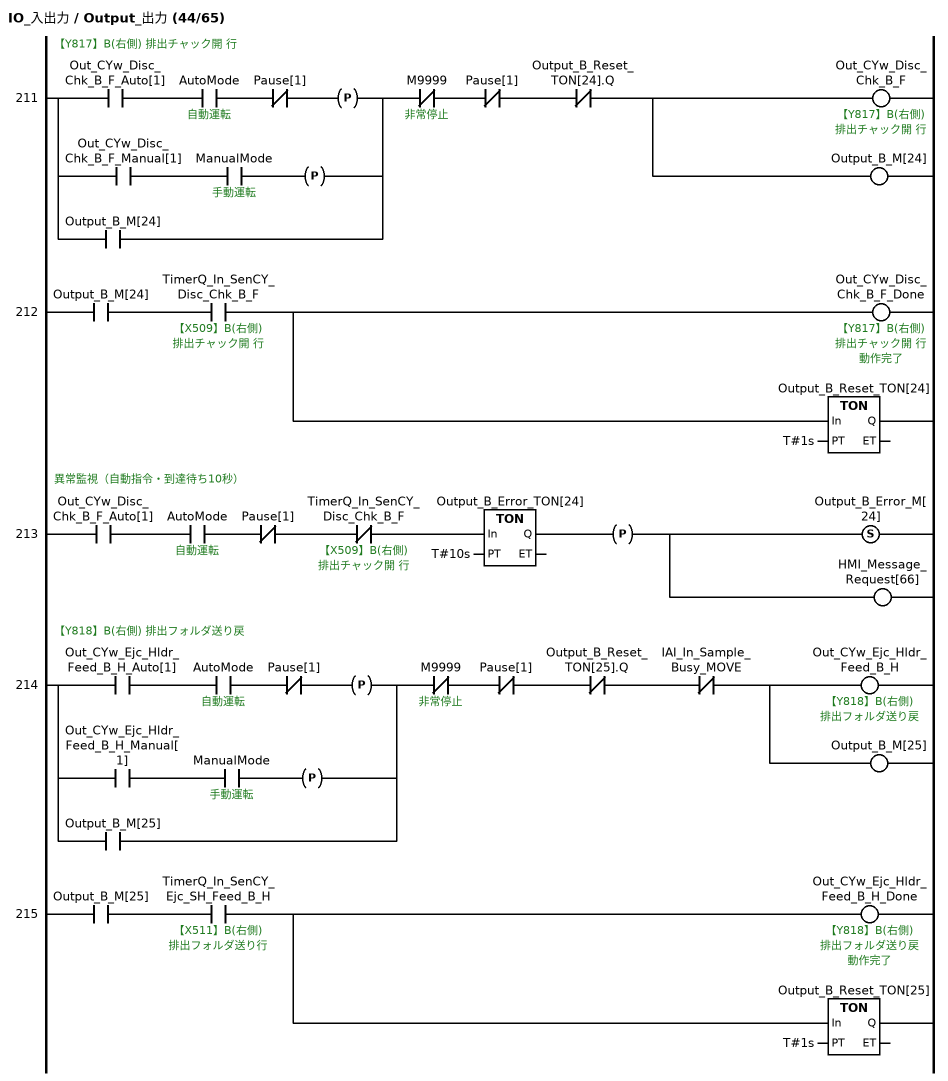
(* [picture p187: IO_入出力 / Output_出力, rungs 211-215] *)
(* Rung 211: 【Y817】B(右側) 排出チャック開 行 *)
_e309(CLK := Out_CYw_Disc_Chk_B_F_Auto[1] AND AutoMode AND NOT Pause[1]);
_e310(CLK := Out_CYw_Disc_Chk_B_F_Manual[1] AND ManualMode);
_p311 := (_e309.Q OR _e310.Q OR Output_B_M[24]) AND NOT M9999 AND NOT Pause[1] AND NOT Output_B_Reset_TON[24].Q;
Out_CYw_Disc_Chk_B_F := _p311;
Output_B_M[24] := _p311;
(* Rung 212 *)
Out_CYw_Disc_Chk_B_F_Done := Output_B_M[24] AND TimerQ_In_SenCY_Disc_Chk_B_F;
Output_B_Reset_TON[24](In := Output_B_M[24] AND TimerQ_In_SenCY_Disc_Chk_B_F, PT := T#1s);
(* Rung 213: 異常監視（自動指令・到達待ち10秒） *)
Output_B_Error_TON[24](In := Out_CYw_Disc_Chk_B_F_Auto[1] AND AutoMode AND NOT Pause[1] AND NOT TimerQ_In_SenCY_Disc_Chk_B_F, PT := T#10s);
_e312(CLK := Output_B_Error_TON[24].Q);
IF _e312.Q THEN Output_B_Error_M[24] := TRUE; END_IF;
HMI_Message_Request[66] := _e312.Q;
(* Rung 214: 【Y818】B(右側) 排出フォルダ送り戻 *)
_e313(CLK := Out_CYw_Ejc_Hldr_Feed_B_H_Auto[1] AND AutoMode AND NOT Pause[1]);
_e314(CLK := Out_CYw_Ejc_Hldr_Feed_B_H_Manual[1] AND ManualMode);
_p315 := (_e313.Q OR _e314.Q OR Output_B_M[25]) AND NOT M9999 AND NOT Pause[1] AND NOT Output_B_Reset_TON[25].Q AND NOT IAI_In_Sample_Busy_MOVE;
Out_CYw_Ejc_Hldr_Feed_B_H := _p315;
Output_B_M[25] := _p315;
(* Rung 215 *)
_p316 := Output_B_M[25] AND TimerQ_In_SenCY_Ejc_SH_Feed_B_H;
Out_CYw_Ejc_Hldr_Feed_B_H_Done := _p316;
Output_B_Reset_TON[25](In := _p316, PT := T#1s);

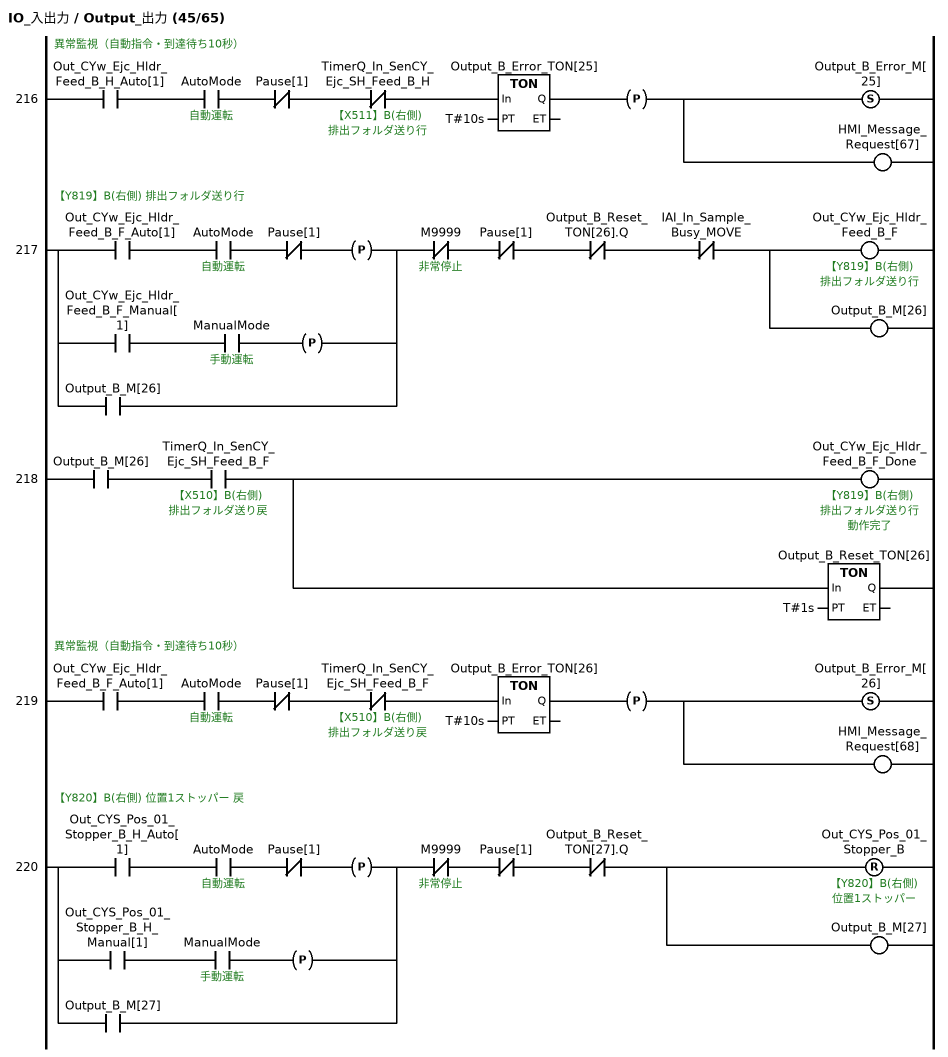
(* Rung 216: 異常監視（自動指令・到達待ち10秒） *)
Output_B_Error_TON[25](In := Out_CYw_Ejc_Hldr_Feed_B_H_Auto[1] AND AutoMode AND NOT Pause[1] AND NOT TimerQ_In_SenCY_Ejc_SH_Feed_B_H, PT := T#10s);
_e317(CLK := Output_B_Error_TON[25].Q);
IF _e317.Q THEN Output_B_Error_M[25] := TRUE; END_IF;
HMI_Message_Request[67] := _e317.Q;
(* Rung 217: 【Y819】B(右側) 排出フォルダ送り行 *)
_e318(CLK := Out_CYw_Ejc_Hldr_Feed_B_F_Auto[1] AND AutoMode AND NOT Pause[1]);
_e319(CLK := Out_CYw_Ejc_Hldr_Feed_B_F_Manual[1] AND ManualMode);
_p320 := (_e318.Q OR _e319.Q OR Output_B_M[26]) AND NOT M9999 AND NOT Pause[1] AND NOT Output_B_Reset_TON[26].Q AND NOT IAI_In_Sample_Busy_MOVE;
Out_CYw_Ejc_Hldr_Feed_B_F := _p320;
Output_B_M[26] := _p320;
(* Rung 218 *)
_p321 := Output_B_M[26] AND TimerQ_In_SenCY_Ejc_SH_Feed_B_F;
Out_CYw_Ejc_Hldr_Feed_B_F_Done := _p321;
Output_B_Reset_TON[26](In := _p321, PT := T#1s);
(* Rung 219: 異常監視（自動指令・到達待ち10秒） *)
Output_B_Error_TON[26](In := Out_CYw_Ejc_Hldr_Feed_B_F_Auto[1] AND AutoMode AND NOT Pause[1] AND NOT TimerQ_In_SenCY_Ejc_SH_Feed_B_F, PT := T#10s);
_e322(CLK := Output_B_Error_TON[26].Q);
IF _e322.Q THEN Output_B_Error_M[26] := TRUE; END_IF;
HMI_Message_Request[68] := _e322.Q;
(* Rung 220: 【Y820】B(右側) 位置1ストッパー 戻 *)
_e323(CLK := Out_CYS_Pos_01_Stopper_B_H_Auto[1] AND AutoMode AND NOT Pause[1]);
_e324(CLK := Out_CYS_Pos_01_Stopper_B_H_Manual[1] AND ManualMode);
_p325 := (_e323.Q OR _e324.Q OR Output_B_M[27]) AND NOT M9999 AND NOT Pause[1] AND NOT Output_B_Reset_TON[27].Q;
IF _p325 THEN Out_CYS_Pos_01_Stopper_B := FALSE; END_IF;
Output_B_M[27] := _p325;

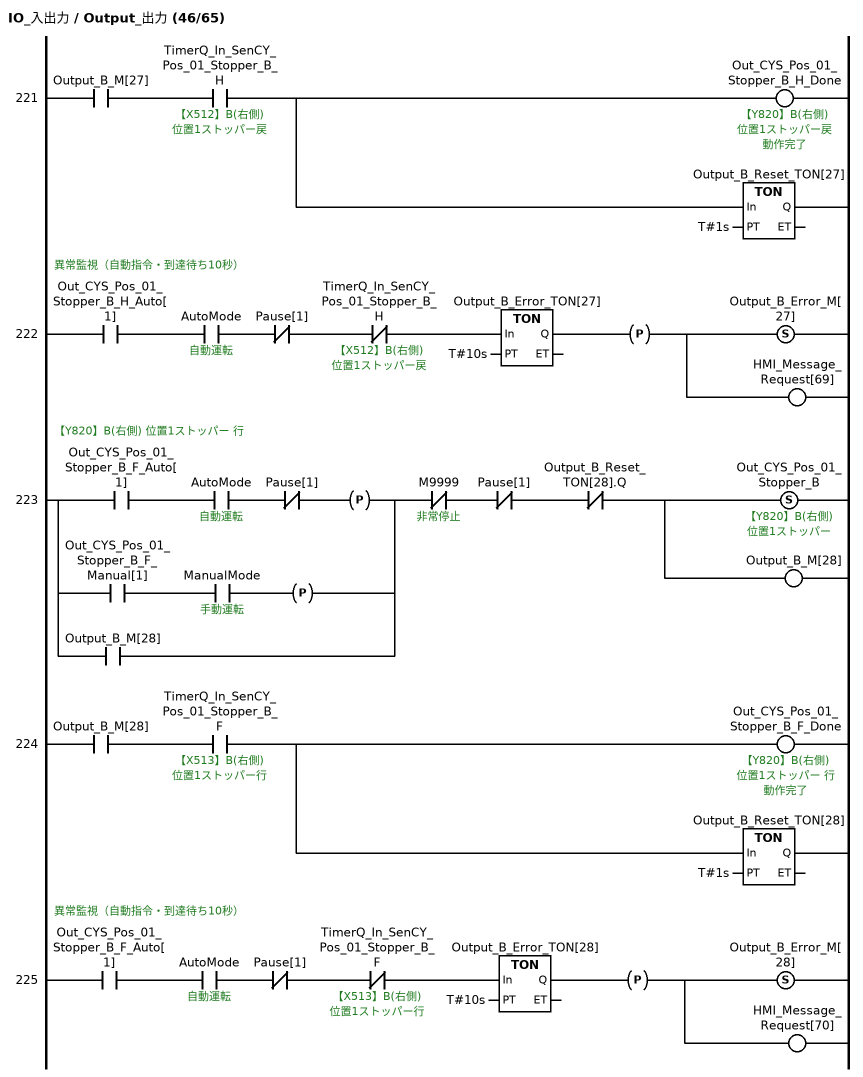
(* Rung 221 *)
_p326 := Output_B_M[27] AND TimerQ_In_SenCY_Pos_01_Stopper_B_H;
Out_CYS_Pos_01_Stopper_B_H_Done := _p326;
Output_B_Reset_TON[27](In := _p326, PT := T#1s);
(* Rung 222: 異常監視（自動指令・到達待ち10秒） *)
Output_B_Error_TON[27](In := Out_CYS_Pos_01_Stopper_B_H_Auto[1] AND AutoMode AND NOT Pause[1] AND NOT TimerQ_In_SenCY_Pos_01_Stopper_B_H, PT := T#10s);
_e327(CLK := Output_B_Error_TON[27].Q);
IF _e327.Q THEN Output_B_Error_M[27] := TRUE; END_IF;
HMI_Message_Request[69] := _e327.Q;
(* Rung 223: 【Y820】B(右側) 位置1ストッパー 行 *)
_e328(CLK := Out_CYS_Pos_01_Stopper_B_F_Auto[1] AND AutoMode AND NOT Pause[1]);
_e329(CLK := Out_CYS_Pos_01_Stopper_B_F_Manual[1] AND ManualMode);
_p330 := (_e328.Q OR _e329.Q OR Output_B_M[28]) AND NOT M9999 AND NOT Pause[1] AND NOT Output_B_Reset_TON[28].Q;
IF _p330 THEN Out_CYS_Pos_01_Stopper_B := TRUE; END_IF;
Output_B_M[28] := _p330;
(* Rung 224 *)
_p331 := Output_B_M[28] AND TimerQ_In_SenCY_Pos_01_Stopper_B_F;
Out_CYS_Pos_01_Stopper_B_F_Done := _p331;
Output_B_Reset_TON[28](In := _p331, PT := T#1s);
(* Rung 225: 異常監視（自動指令・到達待ち10秒） *)
Output_B_Error_TON[28](In := Out_CYS_Pos_01_Stopper_B_F_Auto[1] AND AutoMode AND NOT Pause[1] AND NOT TimerQ_In_SenCY_Pos_01_Stopper_B_F, PT := T#10s);
_e332(CLK := Output_B_Error_TON[28].Q);
IF _e332.Q THEN Output_B_Error_M[28] := TRUE; END_IF;
HMI_Message_Request[70] := _e332.Q;

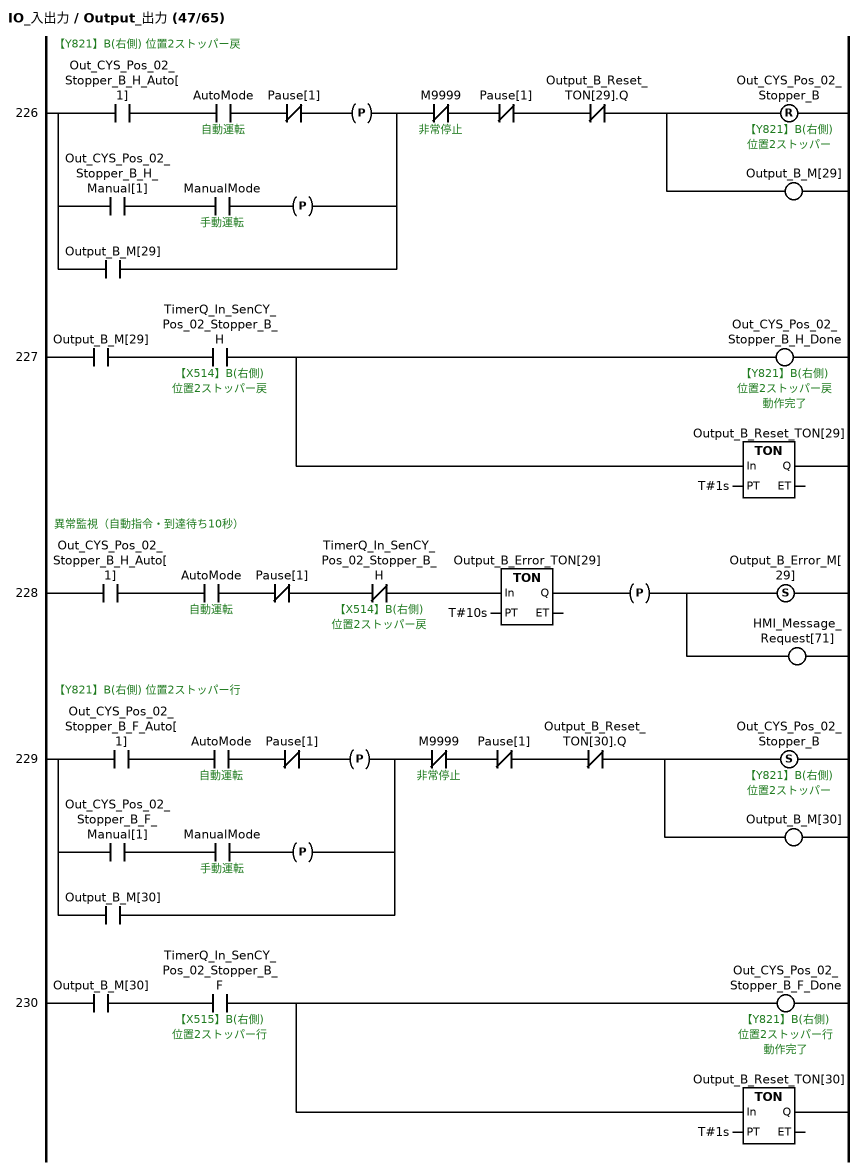
(* Rung 226: 【Y821】B(右側) 位置2ストッパー戻 *)
_e333(CLK := Out_CYS_Pos_02_Stopper_B_H_Auto[1] AND AutoMode AND NOT Pause[1]);
_e334(CLK := Out_CYS_Pos_02_Stopper_B_H_Manual[1] AND ManualMode);
_p335 := (_e333.Q OR _e334.Q OR Output_B_M[29]) AND NOT M9999 AND NOT Pause[1] AND NOT Output_B_Reset_TON[29].Q;
IF _p335 THEN Out_CYS_Pos_02_Stopper_B := FALSE; END_IF;
Output_B_M[29] := _p335;
(* Rung 227 *)
_p336 := Output_B_M[29] AND TimerQ_In_SenCY_Pos_02_Stopper_B_H;
Out_CYS_Pos_02_Stopper_B_H_Done := _p336;
Output_B_Reset_TON[29](In := _p336, PT := T#1s);
(* Rung 228: 異常監視（自動指令・到達待ち10秒） *)
Output_B_Error_TON[29](In := Out_CYS_Pos_02_Stopper_B_H_Auto[1] AND AutoMode AND NOT Pause[1] AND NOT TimerQ_In_SenCY_Pos_02_Stopper_B_H, PT := T#10s);
_e337(CLK := Output_B_Error_TON[29].Q);
IF _e337.Q THEN Output_B_Error_M[29] := TRUE; END_IF;
HMI_Message_Request[71] := _e337.Q;
(* Rung 229: 【Y821】B(右側) 位置2ストッパー行 *)
_e338(CLK := Out_CYS_Pos_02_Stopper_B_F_Auto[1] AND AutoMode AND NOT Pause[1]);
_e339(CLK := Out_CYS_Pos_02_Stopper_B_F_Manual[1] AND ManualMode);
_p340 := (_e338.Q OR _e339.Q OR Output_B_M[30]) AND NOT M9999 AND NOT Pause[1] AND NOT Output_B_Reset_TON[30].Q;
IF _p340 THEN Out_CYS_Pos_02_Stopper_B := TRUE; END_IF;
Output_B_M[30] := _p340;
(* Rung 230 *)
_p341 := Output_B_M[30] AND TimerQ_In_SenCY_Pos_02_Stopper_B_F;
Out_CYS_Pos_02_Stopper_B_F_Done := _p341;
Output_B_Reset_TON[30](In := _p341, PT := T#1s);

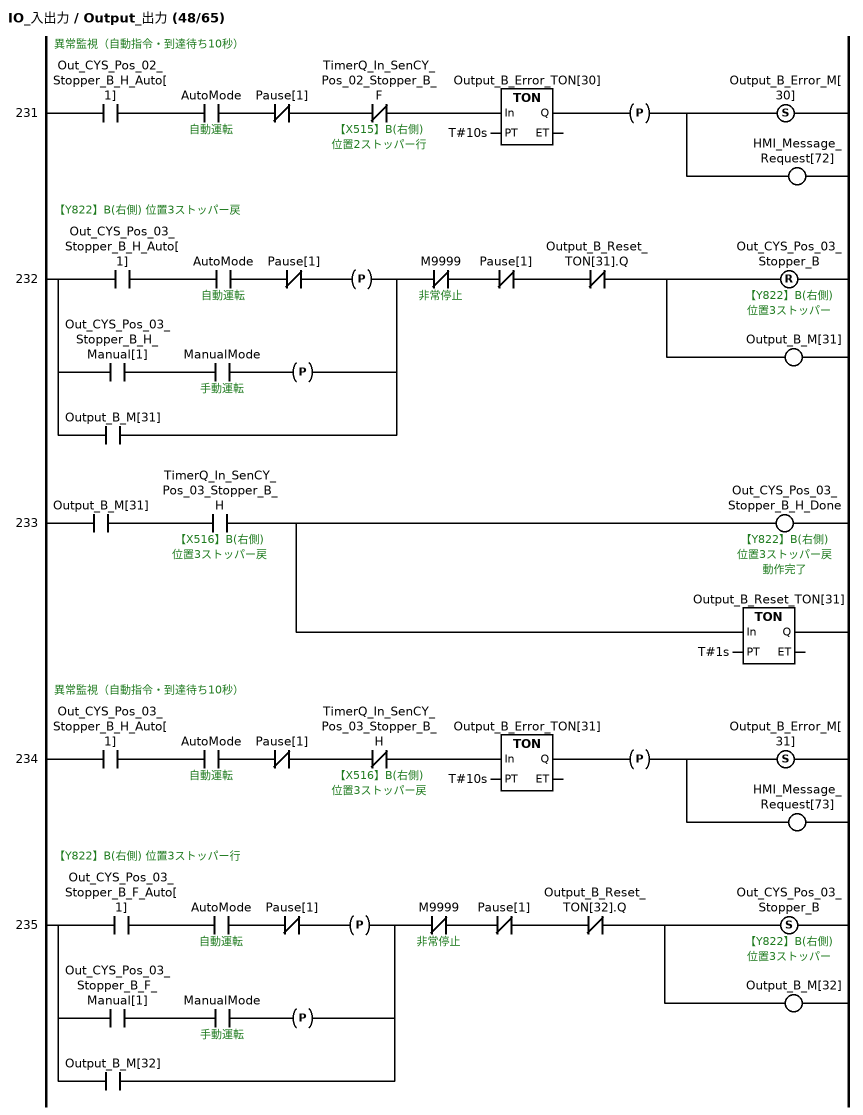
(* Rung 231: 異常監視（自動指令・到達待ち10秒） *)
Output_B_Error_TON[30](In := Out_CYS_Pos_02_Stopper_B_H_Auto[1] AND AutoMode AND NOT Pause[1] AND NOT TimerQ_In_SenCY_Pos_02_Stopper_B_F, PT := T#10s);
_e342(CLK := Output_B_Error_TON[30].Q);
IF _e342.Q THEN Output_B_Error_M[30] := TRUE; END_IF;
HMI_Message_Request[72] := _e342.Q;
(* Rung 232: 【Y822】B(右側) 位置3ストッパー戻 *)
_e343(CLK := Out_CYS_Pos_03_Stopper_B_H_Auto[1] AND AutoMode AND NOT Pause[1]);
_e344(CLK := Out_CYS_Pos_03_Stopper_B_H_Manual[1] AND ManualMode);
_p345 := (_e343.Q OR _e344.Q OR Output_B_M[31]) AND NOT M9999 AND NOT Pause[1] AND NOT Output_B_Reset_TON[31].Q;
IF _p345 THEN Out_CYS_Pos_03_Stopper_B := FALSE; END_IF;
Output_B_M[31] := _p345;
(* Rung 233 *)
_p346 := Output_B_M[31] AND TimerQ_In_SenCY_Pos_03_Stopper_B_H;
Out_CYS_Pos_03_Stopper_B_H_Done := _p346;
Output_B_Reset_TON[31](In := _p346, PT := T#1s);
(* Rung 234: 異常監視（自動指令・到達待ち10秒） *)
Output_B_Error_TON[31](In := Out_CYS_Pos_03_Stopper_B_H_Auto[1] AND AutoMode AND NOT Pause[1] AND NOT TimerQ_In_SenCY_Pos_03_Stopper_B_H, PT := T#10s);
_e347(CLK := Output_B_Error_TON[31].Q);
IF _e347.Q THEN Output_B_Error_M[31] := TRUE; END_IF;
HMI_Message_Request[73] := _e347.Q;
(* Rung 235: 【Y822】B(右側) 位置3ストッパー行 *)
_e348(CLK := Out_CYS_Pos_03_Stopper_B_F_Auto[1] AND AutoMode AND NOT Pause[1]);
_e349(CLK := Out_CYS_Pos_03_Stopper_B_F_Manual[1] AND ManualMode);
_p350 := (_e348.Q OR _e349.Q OR Output_B_M[32]) AND NOT M9999 AND NOT Pause[1] AND NOT Output_B_Reset_TON[32].Q;
IF _p350 THEN Out_CYS_Pos_03_Stopper_B := TRUE; END_IF;
Output_B_M[32] := _p350;

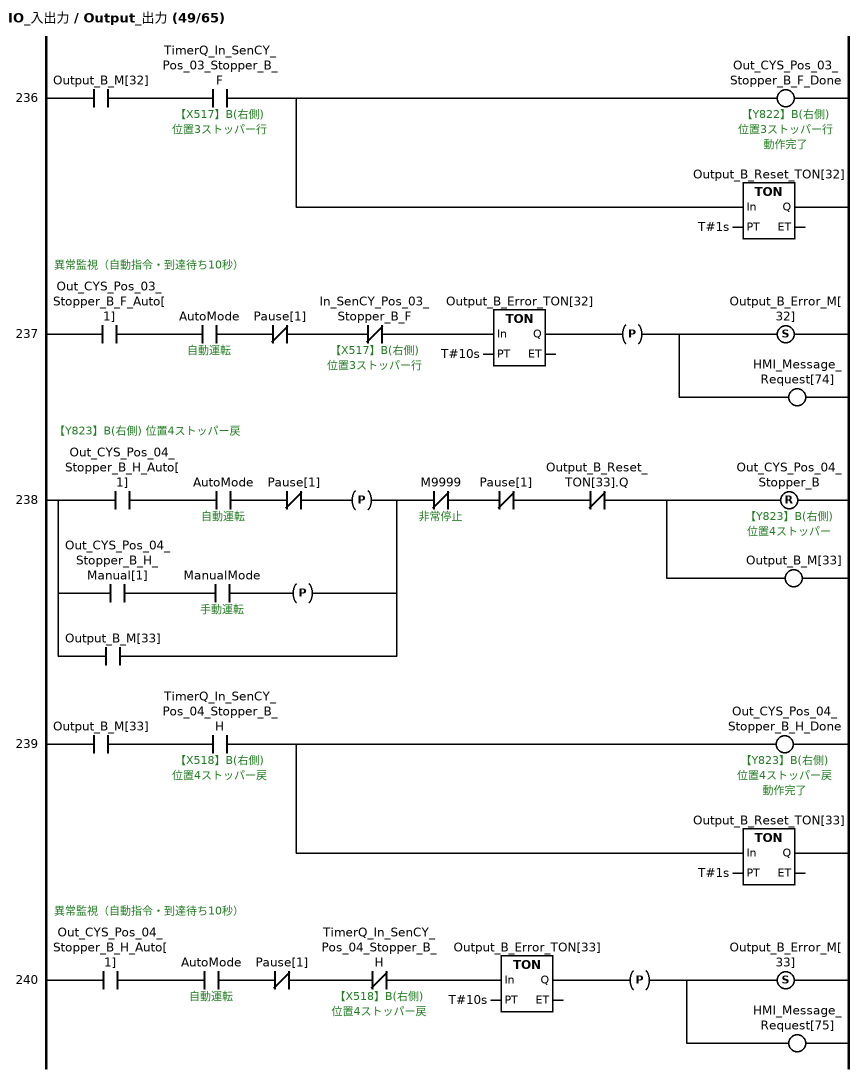
(* Rung 236 *)
_p351 := Output_B_M[32] AND TimerQ_In_SenCY_Pos_03_Stopper_B_F;
Out_CYS_Pos_03_Stopper_B_F_Done := _p351;
Output_B_Reset_TON[32](In := _p351, PT := T#1s);
(* Rung 237: 異常監視（自動指令・到達待ち10秒） *)
Output_B_Error_TON[32](In := Out_CYS_Pos_03_Stopper_B_F_Auto[1] AND AutoMode AND NOT Pause[1] AND NOT In_SenCY_Pos_03_Stopper_B_F, PT := T#10s);
_e352(CLK := Output_B_Error_TON[32].Q);
IF _e352.Q THEN Output_B_Error_M[32] := TRUE; END_IF;
HMI_Message_Request[74] := _e352.Q;
(* Rung 238: 【Y823】B(右側) 位置4ストッパー戻 *)
_e353(CLK := Out_CYS_Pos_04_Stopper_B_H_Auto[1] AND AutoMode AND NOT Pause[1]);
_e354(CLK := Out_CYS_Pos_04_Stopper_B_H_Manual[1] AND ManualMode);
_p355 := (_e353.Q OR _e354.Q OR Output_B_M[33]) AND NOT M9999 AND NOT Pause[1] AND NOT Output_B_Reset_TON[33].Q;
IF _p355 THEN Out_CYS_Pos_04_Stopper_B := FALSE; END_IF;
Output_B_M[33] := _p355;
(* Rung 239 *)
_p356 := Output_B_M[33] AND TimerQ_In_SenCY_Pos_04_Stopper_B_H;
Out_CYS_Pos_04_Stopper_B_H_Done := _p356;
Output_B_Reset_TON[33](In := _p356, PT := T#1s);
(* Rung 240: 異常監視（自動指令・到達待ち10秒） *)
Output_B_Error_TON[33](In := Out_CYS_Pos_04_Stopper_B_H_Auto[1] AND AutoMode AND NOT Pause[1] AND NOT TimerQ_In_SenCY_Pos_04_Stopper_B_H, PT := T#10s);
_e357(CLK := Output_B_Error_TON[33].Q);
IF _e357.Q THEN Output_B_Error_M[33] := TRUE; END_IF;
HMI_Message_Request[75] := _e357.Q;

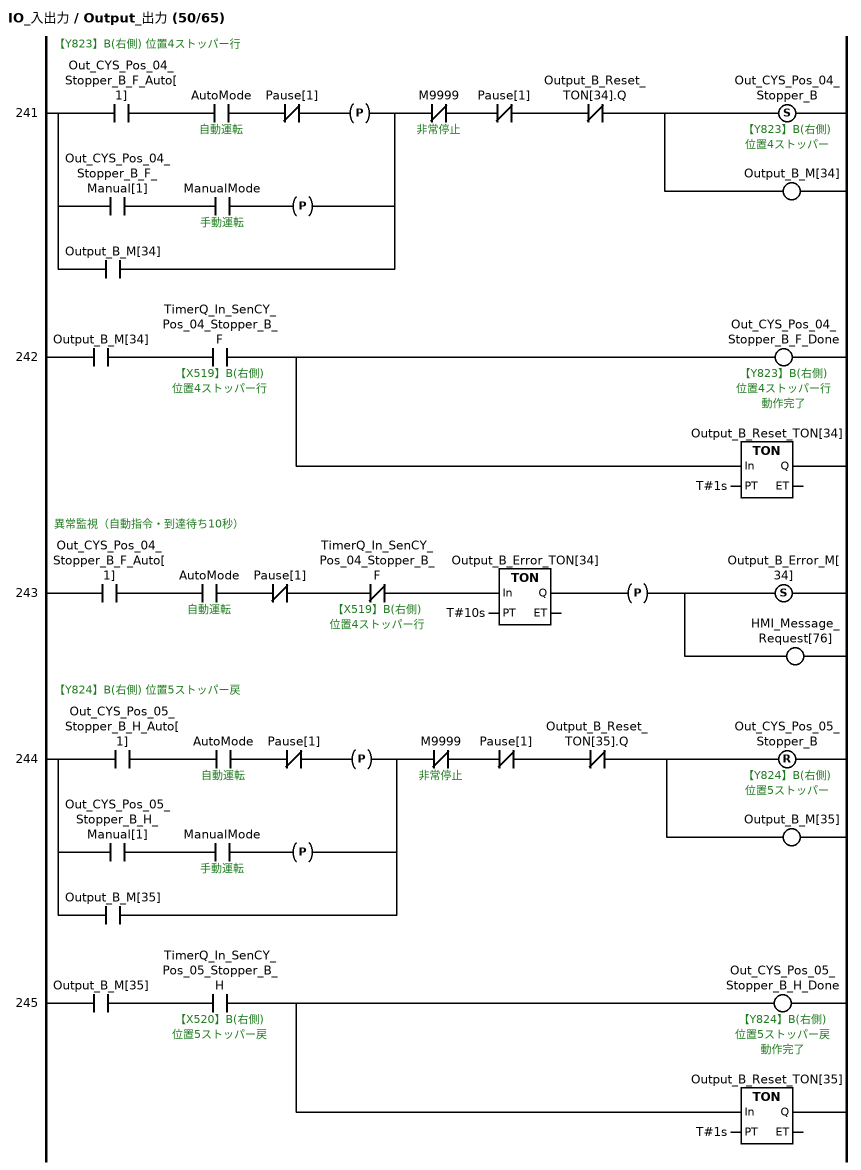
(* Rung 241: 【Y823】B(右側) 位置4ストッパー行 *)
_e358(CLK := Out_CYS_Pos_04_Stopper_B_F_Auto[1] AND AutoMode AND NOT Pause[1]);
_e359(CLK := Out_CYS_Pos_04_Stopper_B_F_Manual[1] AND ManualMode);
_p360 := (_e358.Q OR _e359.Q OR Output_B_M[34]) AND NOT M9999 AND NOT Pause[1] AND NOT Output_B_Reset_TON[34].Q;
IF _p360 THEN Out_CYS_Pos_04_Stopper_B := TRUE; END_IF;
Output_B_M[34] := _p360;
(* Rung 242 *)
_p361 := Output_B_M[34] AND TimerQ_In_SenCY_Pos_04_Stopper_B_F;
Out_CYS_Pos_04_Stopper_B_F_Done := _p361;
Output_B_Reset_TON[34](In := _p361, PT := T#1s);
(* Rung 243: 異常監視（自動指令・到達待ち10秒） *)
Output_B_Error_TON[34](In := Out_CYS_Pos_04_Stopper_B_F_Auto[1] AND AutoMode AND NOT Pause[1] AND NOT TimerQ_In_SenCY_Pos_04_Stopper_B_F, PT := T#10s);
_e362(CLK := Output_B_Error_TON[34].Q);
IF _e362.Q THEN Output_B_Error_M[34] := TRUE; END_IF;
HMI_Message_Request[76] := _e362.Q;
(* Rung 244: 【Y824】B(右側) 位置5ストッパー戻 *)
_e363(CLK := Out_CYS_Pos_05_Stopper_B_H_Auto[1] AND AutoMode AND NOT Pause[1]);
_e364(CLK := Out_CYS_Pos_05_Stopper_B_H_Manual[1] AND ManualMode);
_p365 := (_e363.Q OR _e364.Q OR Output_B_M[35]) AND NOT M9999 AND NOT Pause[1] AND NOT Output_B_Reset_TON[35].Q;
IF _p365 THEN Out_CYS_Pos_05_Stopper_B := FALSE; END_IF;
Output_B_M[35] := _p365;
(* Rung 245 *)
_p366 := Output_B_M[35] AND TimerQ_In_SenCY_Pos_05_Stopper_B_H;
Out_CYS_Pos_05_Stopper_B_H_Done := _p366;
Output_B_Reset_TON[35](In := _p366, PT := T#1s);

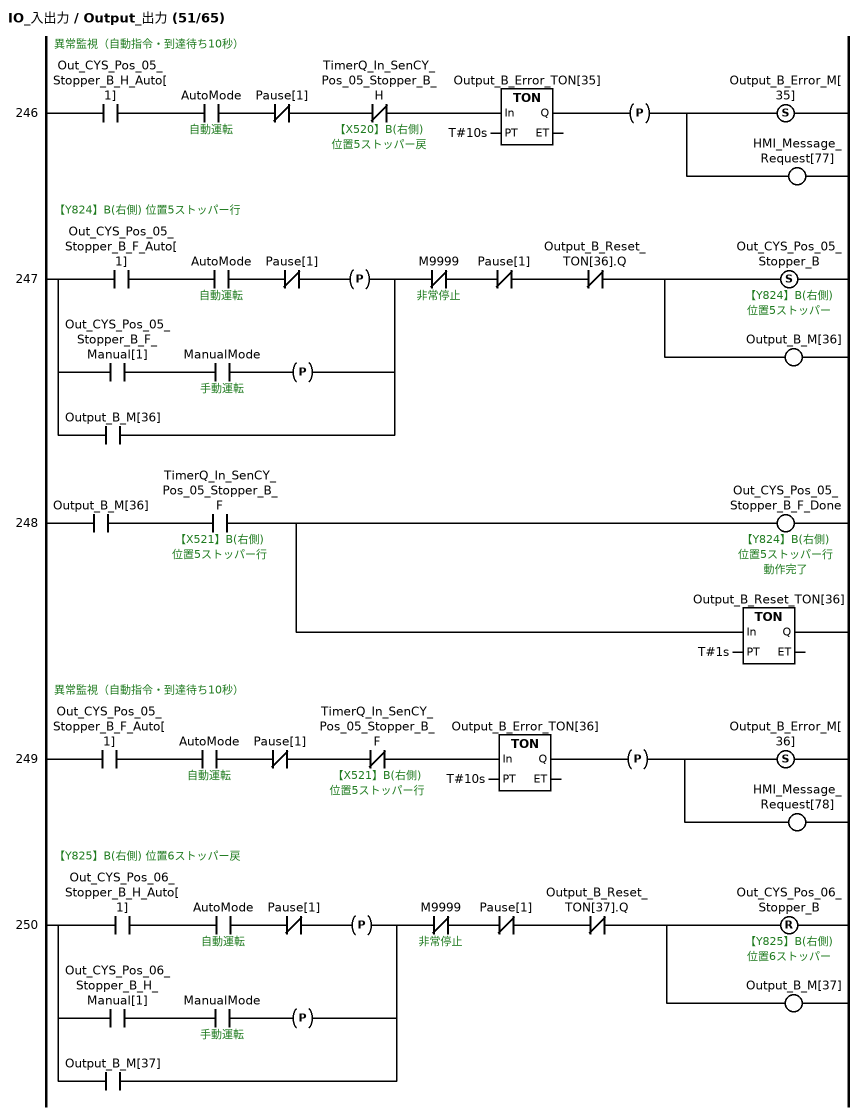
(* Rung 246: 異常監視（自動指令・到達待ち10秒） *)
Output_B_Error_TON[35](In := Out_CYS_Pos_05_Stopper_B_H_Auto[1] AND AutoMode AND NOT Pause[1] AND NOT TimerQ_In_SenCY_Pos_05_Stopper_B_H, PT := T#10s);
_e367(CLK := Output_B_Error_TON[35].Q);
IF _e367.Q THEN Output_B_Error_M[35] := TRUE; END_IF;
HMI_Message_Request[77] := _e367.Q;
(* Rung 247: 【Y824】B(右側) 位置5ストッパー行 *)
_e368(CLK := Out_CYS_Pos_05_Stopper_B_F_Auto[1] AND AutoMode AND NOT Pause[1]);
_e369(CLK := Out_CYS_Pos_05_Stopper_B_F_Manual[1] AND ManualMode);
_p370 := (_e368.Q OR _e369.Q OR Output_B_M[36]) AND NOT M9999 AND NOT Pause[1] AND NOT Output_B_Reset_TON[36].Q;
IF _p370 THEN Out_CYS_Pos_05_Stopper_B := TRUE; END_IF;
Output_B_M[36] := _p370;
(* Rung 248 *)
_p371 := Output_B_M[36] AND TimerQ_In_SenCY_Pos_05_Stopper_B_F;
Out_CYS_Pos_05_Stopper_B_F_Done := _p371;
Output_B_Reset_TON[36](In := _p371, PT := T#1s);
(* Rung 249: 異常監視（自動指令・到達待ち10秒） *)
Output_B_Error_TON[36](In := Out_CYS_Pos_05_Stopper_B_F_Auto[1] AND AutoMode AND NOT Pause[1] AND NOT TimerQ_In_SenCY_Pos_05_Stopper_B_F, PT := T#10s);
_e372(CLK := Output_B_Error_TON[36].Q);
IF _e372.Q THEN Output_B_Error_M[36] := TRUE; END_IF;
HMI_Message_Request[78] := _e372.Q;
(* Rung 250: 【Y825】B(右側) 位置6ストッパー戻 *)
_e373(CLK := Out_CYS_Pos_06_Stopper_B_H_Auto[1] AND AutoMode AND NOT Pause[1]);
_e374(CLK := Out_CYS_Pos_06_Stopper_B_H_Manual[1] AND ManualMode);
_p375 := (_e373.Q OR _e374.Q OR Output_B_M[37]) AND NOT M9999 AND NOT Pause[1] AND NOT Output_B_Reset_TON[37].Q;
IF _p375 THEN Out_CYS_Pos_06_Stopper_B := FALSE; END_IF;
Output_B_M[37] := _p375;

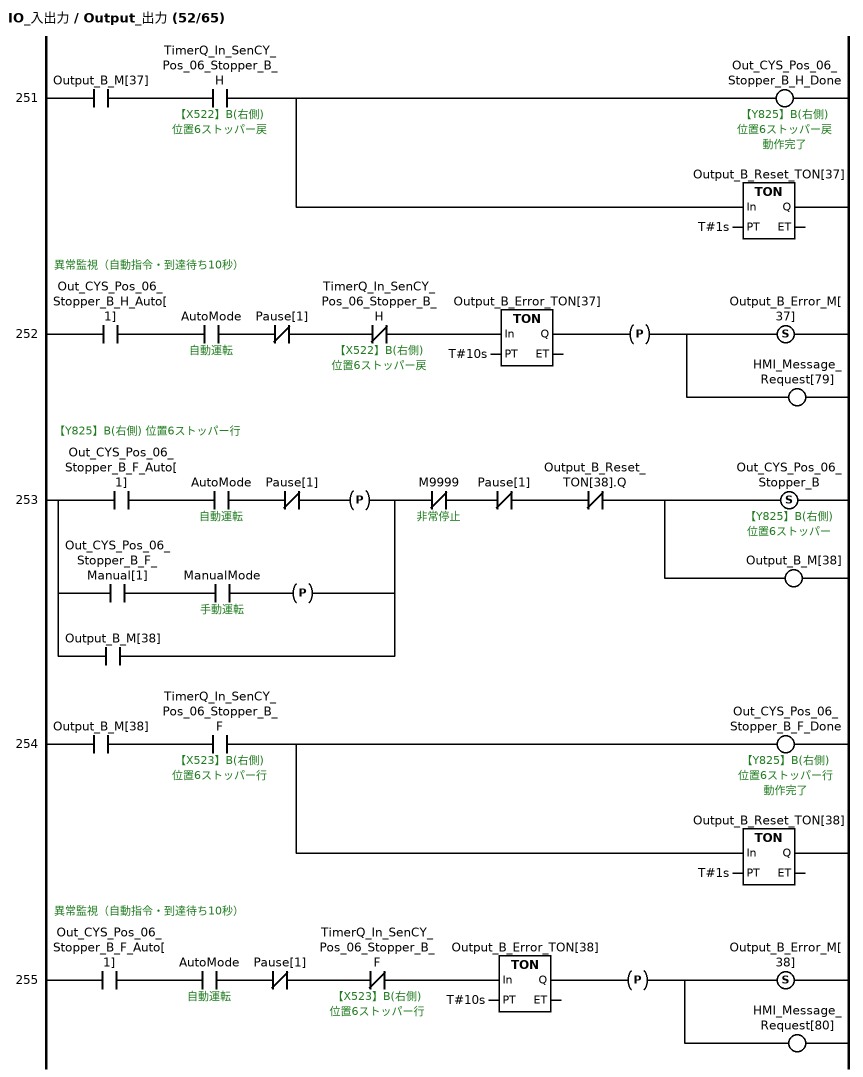
(* Rung 251 *)
_p376 := Output_B_M[37] AND TimerQ_In_SenCY_Pos_06_Stopper_B_H;
Out_CYS_Pos_06_Stopper_B_H_Done := _p376;
Output_B_Reset_TON[37](In := _p376, PT := T#1s);
(* Rung 252: 異常監視（自動指令・到達待ち10秒） *)
Output_B_Error_TON[37](In := Out_CYS_Pos_06_Stopper_B_H_Auto[1] AND AutoMode AND NOT Pause[1] AND NOT TimerQ_In_SenCY_Pos_06_Stopper_B_H, PT := T#10s);
_e377(CLK := Output_B_Error_TON[37].Q);
IF _e377.Q THEN Output_B_Error_M[37] := TRUE; END_IF;
HMI_Message_Request[79] := _e377.Q;
(* Rung 253: 【Y825】B(右側) 位置6ストッパー行 *)
_e378(CLK := Out_CYS_Pos_06_Stopper_B_F_Auto[1] AND AutoMode AND NOT Pause[1]);
_e379(CLK := Out_CYS_Pos_06_Stopper_B_F_Manual[1] AND ManualMode);
_p380 := (_e378.Q OR _e379.Q OR Output_B_M[38]) AND NOT M9999 AND NOT Pause[1] AND NOT Output_B_Reset_TON[38].Q;
IF _p380 THEN Out_CYS_Pos_06_Stopper_B := TRUE; END_IF;
Output_B_M[38] := _p380;
(* Rung 254 *)
_p381 := Output_B_M[38] AND TimerQ_In_SenCY_Pos_06_Stopper_B_F;
Out_CYS_Pos_06_Stopper_B_F_Done := _p381;
Output_B_Reset_TON[38](In := _p381, PT := T#1s);
(* Rung 255: 異常監視（自動指令・到達待ち10秒） *)
Output_B_Error_TON[38](In := Out_CYS_Pos_06_Stopper_B_F_Auto[1] AND AutoMode AND NOT Pause[1] AND NOT TimerQ_In_SenCY_Pos_06_Stopper_B_F, PT := T#10s);
_e382(CLK := Output_B_Error_TON[38].Q);
IF _e382.Q THEN Output_B_Error_M[38] := TRUE; END_IF;
HMI_Message_Request[80] := _e382.Q;

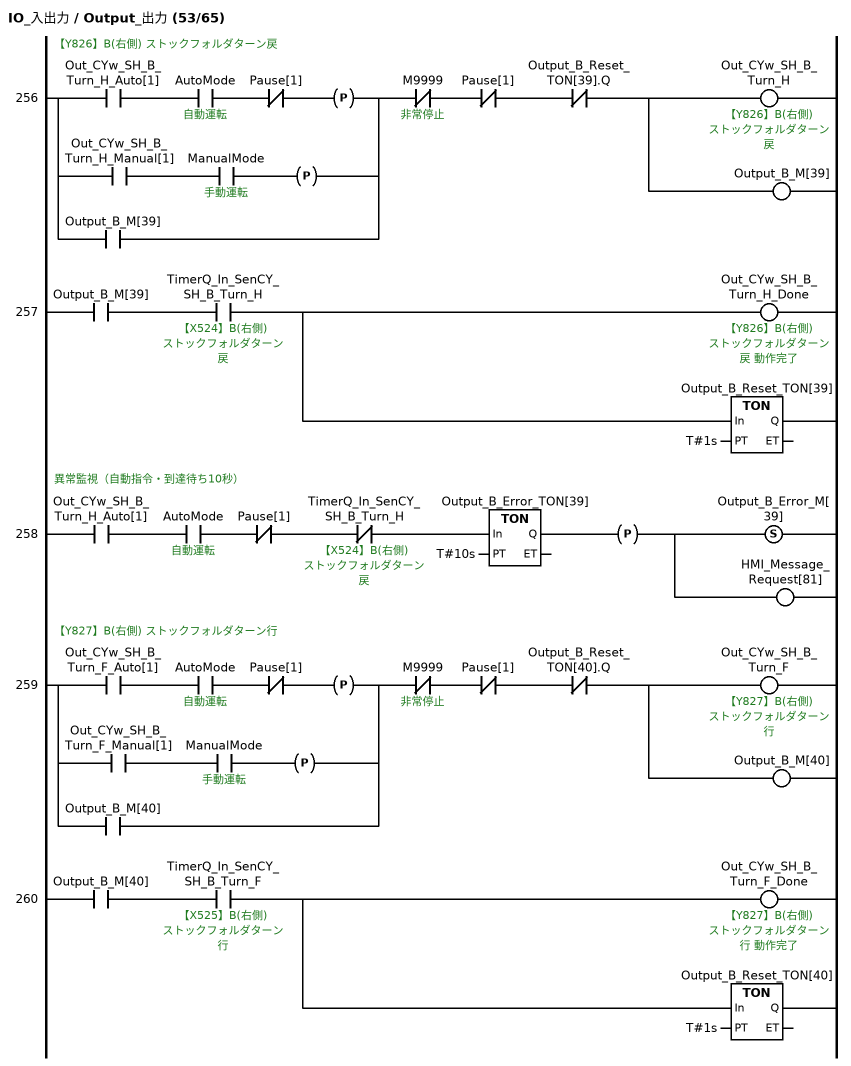
(* Rung 256: 【Y826】B(右側) ストックフォルダターン戻 *)
_e383(CLK := Out_CYw_SH_B_Turn_H_Auto[1] AND AutoMode AND NOT Pause[1]);
_e384(CLK := Out_CYw_SH_B_Turn_H_Manual[1] AND ManualMode);
_p385 := (_e383.Q OR _e384.Q OR Output_B_M[39]) AND NOT M9999 AND NOT Pause[1] AND NOT Output_B_Reset_TON[39].Q;
Out_CYw_SH_B_Turn_H := _p385;
Output_B_M[39] := _p385;
(* Rung 257 *)
Out_CYw_SH_B_Turn_H_Done := Output_B_M[39] AND TimerQ_In_SenCY_SH_B_Turn_H;
Output_B_Reset_TON[39](In := Output_B_M[39] AND TimerQ_In_SenCY_SH_B_Turn_H, PT := T#1s);
(* Rung 258: 異常監視（自動指令・到達待ち10秒） *)
Output_B_Error_TON[39](In := Out_CYw_SH_B_Turn_H_Auto[1] AND AutoMode AND NOT Pause[1] AND NOT TimerQ_In_SenCY_SH_B_Turn_H, PT := T#10s);
_e386(CLK := Output_B_Error_TON[39].Q);
IF _e386.Q THEN Output_B_Error_M[39] := TRUE; END_IF;
HMI_Message_Request[81] := _e386.Q;
(* Rung 259: 【Y827】B(右側) ストックフォルダターン行 *)
_e387(CLK := Out_CYw_SH_B_Turn_F_Auto[1] AND AutoMode AND NOT Pause[1]);
_e388(CLK := Out_CYw_SH_B_Turn_F_Manual[1] AND ManualMode);
_p389 := (_e387.Q OR _e388.Q OR Output_B_M[40]) AND NOT M9999 AND NOT Pause[1] AND NOT Output_B_Reset_TON[40].Q;
Out_CYw_SH_B_Turn_F := _p389;
Output_B_M[40] := _p389;
(* Rung 260 *)
Out_CYw_SH_B_Turn_F_Done := Output_B_M[40] AND TimerQ_In_SenCY_SH_B_Turn_F;
Output_B_Reset_TON[40](In := Output_B_M[40] AND TimerQ_In_SenCY_SH_B_Turn_F, PT := T#1s);

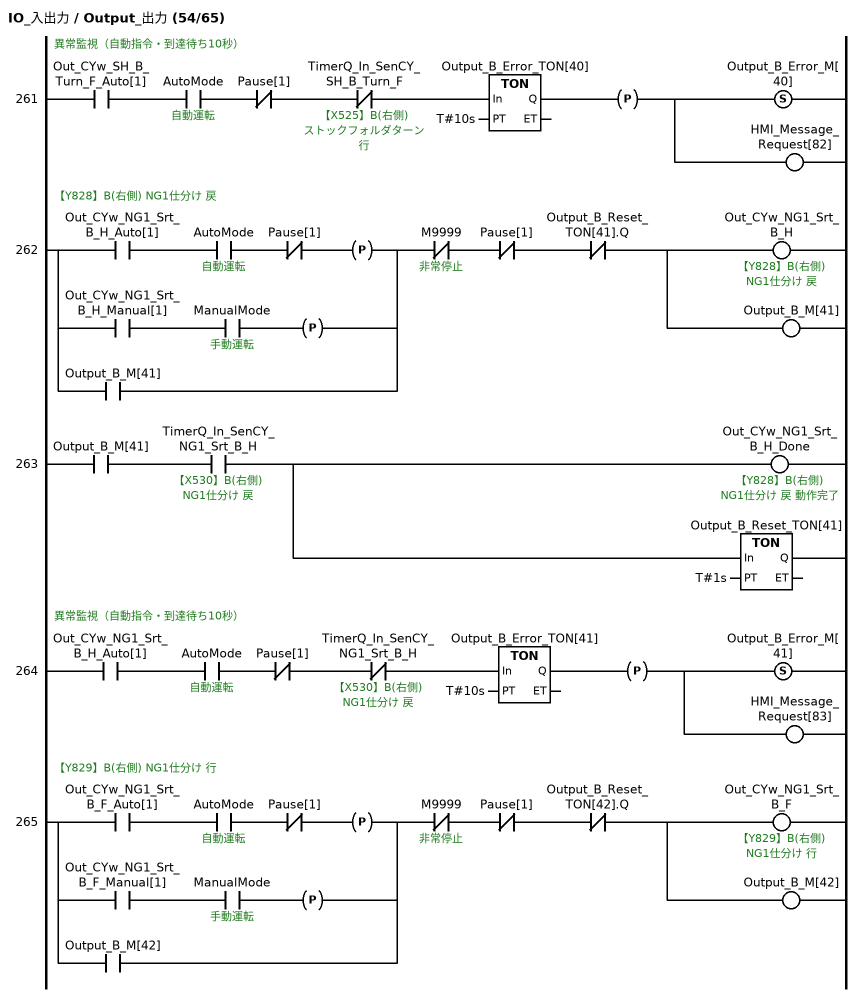
(* Rung 261: 異常監視（自動指令・到達待ち10秒） *)
Output_B_Error_TON[40](In := Out_CYw_SH_B_Turn_F_Auto[1] AND AutoMode AND NOT Pause[1] AND NOT TimerQ_In_SenCY_SH_B_Turn_F, PT := T#10s);
_e390(CLK := Output_B_Error_TON[40].Q);
IF _e390.Q THEN Output_B_Error_M[40] := TRUE; END_IF;
HMI_Message_Request[82] := _e390.Q;
(* Rung 262: 【Y828】B(右側) NG1仕分け 戻 *)
_e391(CLK := Out_CYw_NG1_Srt_B_H_Auto[1] AND AutoMode AND NOT Pause[1]);
_e392(CLK := Out_CYw_NG1_Srt_B_H_Manual[1] AND ManualMode);
_p393 := (_e391.Q OR _e392.Q OR Output_B_M[41]) AND NOT M9999 AND NOT Pause[1] AND NOT Output_B_Reset_TON[41].Q;
Out_CYw_NG1_Srt_B_H := _p393;
Output_B_M[41] := _p393;
(* Rung 263 *)
Out_CYw_NG1_Srt_B_H_Done := Output_B_M[41] AND TimerQ_In_SenCY_NG1_Srt_B_H;
Output_B_Reset_TON[41](In := Output_B_M[41] AND TimerQ_In_SenCY_NG1_Srt_B_H, PT := T#1s);
(* Rung 264: 異常監視（自動指令・到達待ち10秒） *)
Output_B_Error_TON[41](In := Out_CYw_NG1_Srt_B_H_Auto[1] AND AutoMode AND NOT Pause[1] AND NOT TimerQ_In_SenCY_NG1_Srt_B_H, PT := T#10s);
_e394(CLK := Output_B_Error_TON[41].Q);
IF _e394.Q THEN Output_B_Error_M[41] := TRUE; END_IF;
HMI_Message_Request[83] := _e394.Q;
(* Rung 265: 【Y829】B(右側) NG1仕分け 行 *)
_e395(CLK := Out_CYw_NG1_Srt_B_F_Auto[1] AND AutoMode AND NOT Pause[1]);
_e396(CLK := Out_CYw_NG1_Srt_B_F_Manual[1] AND ManualMode);
_p397 := (_e395.Q OR _e396.Q OR Output_B_M[42]) AND NOT M9999 AND NOT Pause[1] AND NOT Output_B_Reset_TON[42].Q;
Out_CYw_NG1_Srt_B_F := _p397;
Output_B_M[42] := _p397;

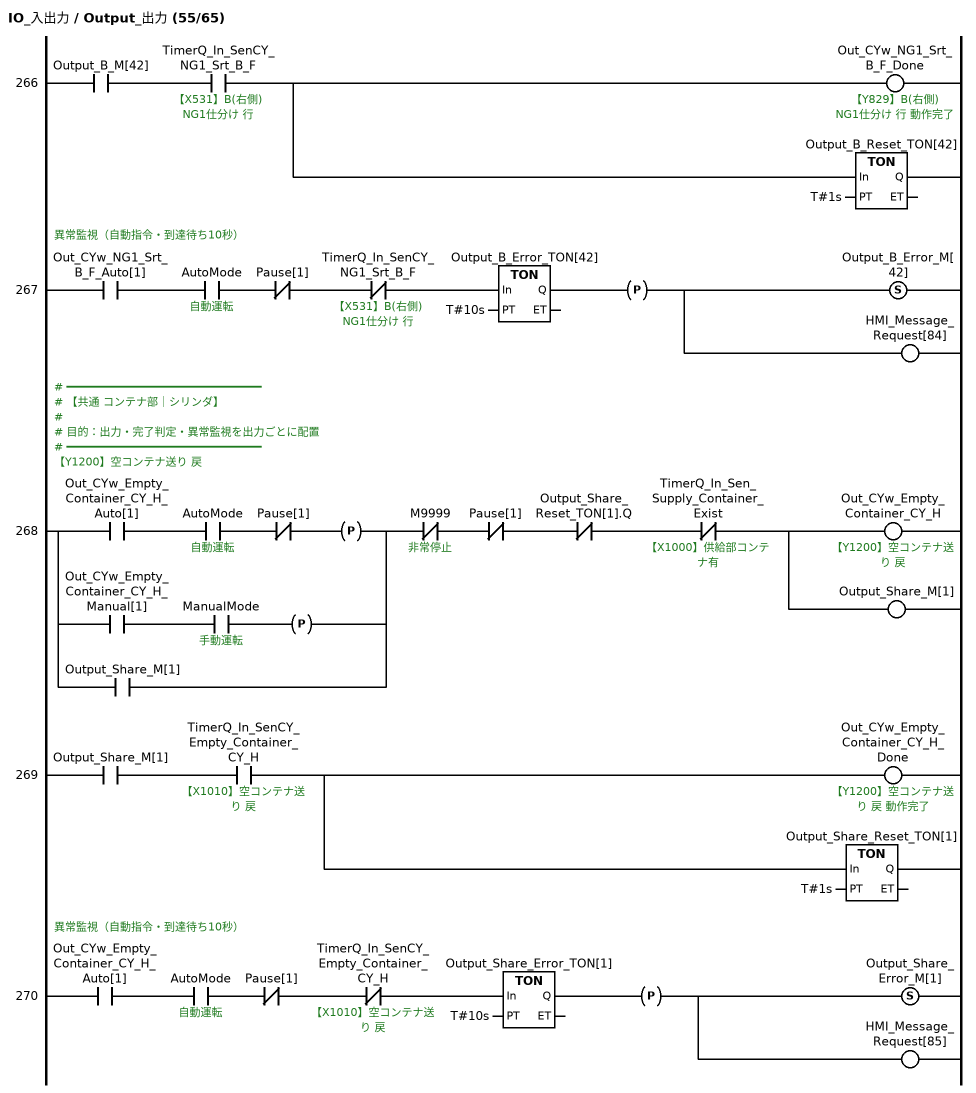
(* Rung 266 *)
Out_CYw_NG1_Srt_B_F_Done := Output_B_M[42] AND TimerQ_In_SenCY_NG1_Srt_B_F;
Output_B_Reset_TON[42](In := Output_B_M[42] AND TimerQ_In_SenCY_NG1_Srt_B_F, PT := T#1s);
(* Rung 267: 異常監視（自動指令・到達待ち10秒） *)
Output_B_Error_TON[42](In := Out_CYw_NG1_Srt_B_F_Auto[1] AND AutoMode AND NOT Pause[1] AND NOT TimerQ_In_SenCY_NG1_Srt_B_F, PT := T#10s);
_e398(CLK := Output_B_Error_TON[42].Q);
IF _e398.Q THEN Output_B_Error_M[42] := TRUE; END_IF;
HMI_Message_Request[84] := _e398.Q;
(* Rung 268: # ━━━━━━━━━━━━━━━━━━━━━━━━━━━━━━ / # 【共通 コンテナ部｜シリンダ】 / # / # 目的：出力・完了判定・異常監視を出力ごとに配置 / # ━━━━━━━━━━━━━━━━━━━━━━━━━━━━━━ / 【Y1200】空コンテナ送り 戻 *)
_e399(CLK := Out_CYw_Empty_Container_CY_H_Auto[1] AND AutoMode AND NOT Pause[1]);
_e400(CLK := Out_CYw_Empty_Container_CY_H_Manual[1] AND ManualMode);
_p401 := (_e399.Q OR _e400.Q OR Output_Share_M[1]) AND NOT M9999 AND NOT Pause[1] AND NOT Output_Share_Reset_TON[1].Q AND NOT TimerQ_In_Sen_Supply_Container_Exist;
Out_CYw_Empty_Container_CY_H := _p401;
Output_Share_M[1] := _p401;
(* Rung 269 *)
_p402 := Output_Share_M[1] AND TimerQ_In_SenCY_Empty_Container_CY_H;
Out_CYw_Empty_Container_CY_H_Done := _p402;
Output_Share_Reset_TON[1](In := _p402, PT := T#1s);
(* Rung 270: 異常監視（自動指令・到達待ち10秒） *)
Output_Share_Error_TON[1](In := Out_CYw_Empty_Container_CY_H_Auto[1] AND AutoMode AND NOT Pause[1] AND NOT TimerQ_In_SenCY_Empty_Container_CY_H, PT := T#10s);
_e403(CLK := Output_Share_Error_TON[1].Q);
IF _e403.Q THEN Output_Share_Error_M[1] := TRUE; END_IF;
HMI_Message_Request[85] := _e403.Q;

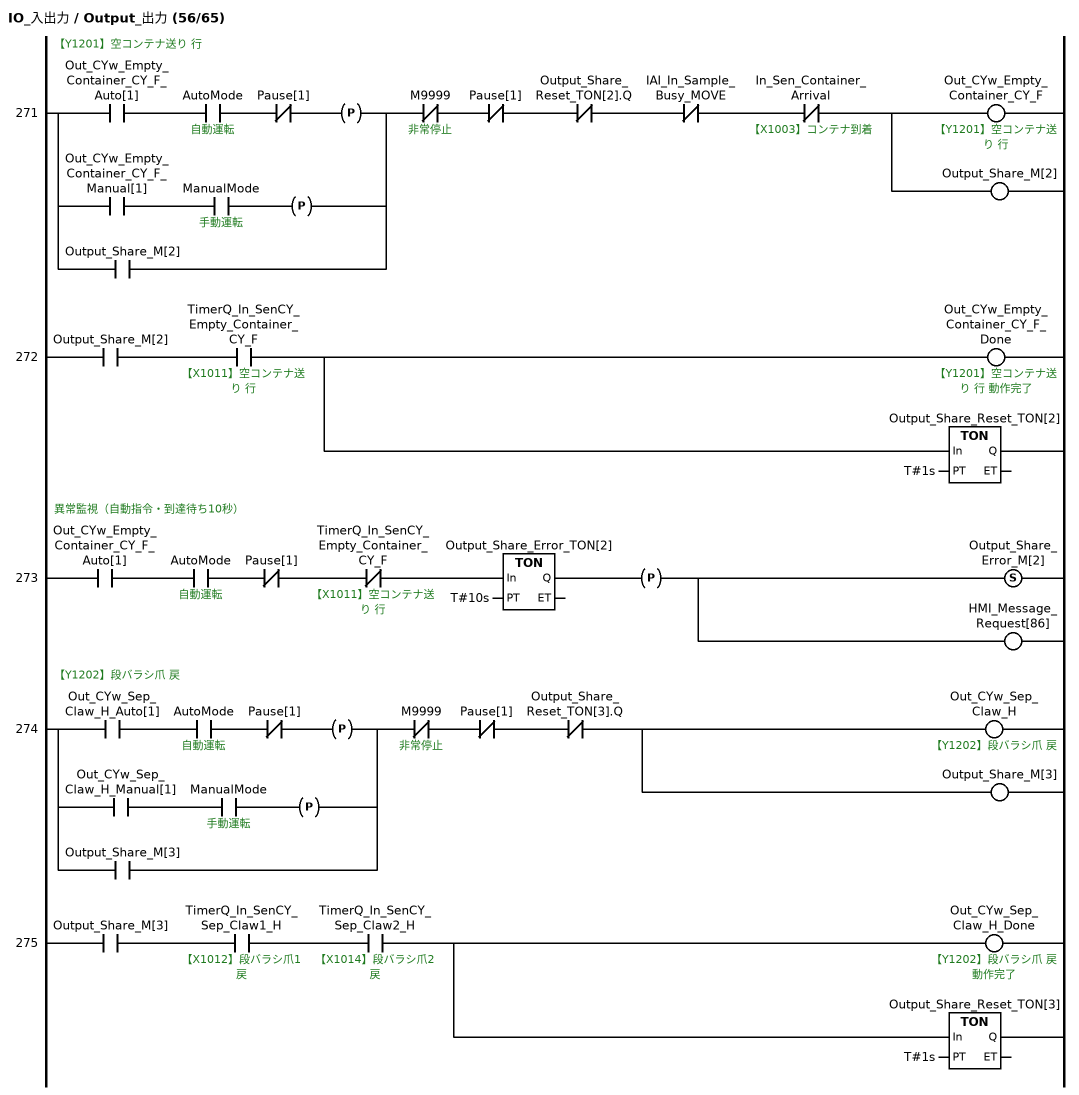
(* Rung 271: 【Y1201】空コンテナ送り 行 *)
_e404(CLK := Out_CYw_Empty_Container_CY_F_Auto[1] AND AutoMode AND NOT Pause[1]);
_e405(CLK := Out_CYw_Empty_Container_CY_F_Manual[1] AND ManualMode);
_p406 := (_e404.Q OR _e405.Q OR Output_Share_M[2]) AND NOT M9999 AND NOT Pause[1] AND NOT Output_Share_Reset_TON[2].Q AND NOT IAI_In_Sample_Busy_MOVE AND NOT In_Sen_Container_Arrival;
Out_CYw_Empty_Container_CY_F := _p406;
Output_Share_M[2] := _p406;
(* Rung 272 *)
_p407 := Output_Share_M[2] AND TimerQ_In_SenCY_Empty_Container_CY_F;
Out_CYw_Empty_Container_CY_F_Done := _p407;
Output_Share_Reset_TON[2](In := _p407, PT := T#1s);
(* Rung 273: 異常監視（自動指令・到達待ち10秒） *)
Output_Share_Error_TON[2](In := Out_CYw_Empty_Container_CY_F_Auto[1] AND AutoMode AND NOT Pause[1] AND NOT TimerQ_In_SenCY_Empty_Container_CY_F, PT := T#10s);
_e408(CLK := Output_Share_Error_TON[2].Q);
IF _e408.Q THEN Output_Share_Error_M[2] := TRUE; END_IF;
HMI_Message_Request[86] := _e408.Q;
(* Rung 274: 【Y1202】段バラシ爪 戻 *)
_e409(CLK := Out_CYw_Sep_Claw_H_Auto[1] AND AutoMode AND NOT Pause[1]);
_e410(CLK := Out_CYw_Sep_Claw_H_Manual[1] AND ManualMode);
_p411 := (_e409.Q OR _e410.Q OR Output_Share_M[3]) AND NOT M9999 AND NOT Pause[1] AND NOT Output_Share_Reset_TON[3].Q;
Out_CYw_Sep_Claw_H := _p411;
Output_Share_M[3] := _p411;
(* Rung 275 *)
_p412 := Output_Share_M[3] AND TimerQ_In_SenCY_Sep_Claw1_H AND TimerQ_In_SenCY_Sep_Claw2_H;
Out_CYw_Sep_Claw_H_Done := _p412;
Output_Share_Reset_TON[3](In := _p412, PT := T#1s);

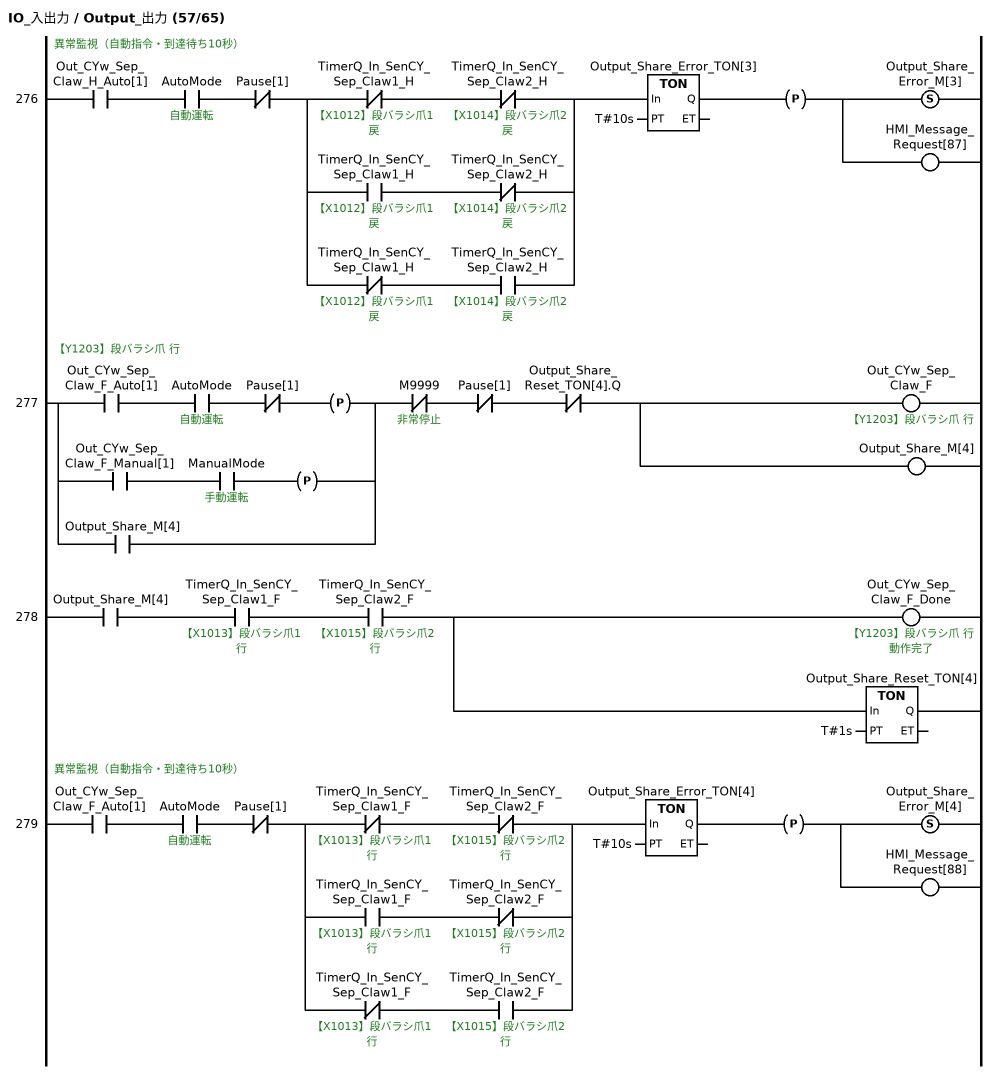
(* Rung 276: 異常監視（自動指令・到達待ち10秒） *)
Output_Share_Error_TON[3](In := Out_CYw_Sep_Claw_H_Auto[1] AND AutoMode AND NOT Pause[1] AND ((NOT TimerQ_In_SenCY_Sep_Claw1_H AND NOT TimerQ_In_SenCY_Sep_Claw2_H) OR (TimerQ_In_SenCY_Sep_Claw1_H AND NOT TimerQ_In_SenCY_Sep_Claw2_H) OR (NOT TimerQ_In_SenCY_Sep_Claw1_H AND TimerQ_In_SenCY_Sep_Claw2_H)), PT := T#10s);
_e413(CLK := Output_Share_Error_TON[3].Q);
IF _e413.Q THEN Output_Share_Error_M[3] := TRUE; END_IF;
HMI_Message_Request[87] := _e413.Q;
(* Rung 277: 【Y1203】段バラシ爪 行 *)
_e414(CLK := Out_CYw_Sep_Claw_F_Auto[1] AND AutoMode AND NOT Pause[1]);
_e415(CLK := Out_CYw_Sep_Claw_F_Manual[1] AND ManualMode);
_p416 := (_e414.Q OR _e415.Q OR Output_Share_M[4]) AND NOT M9999 AND NOT Pause[1] AND NOT Output_Share_Reset_TON[4].Q;
Out_CYw_Sep_Claw_F := _p416;
Output_Share_M[4] := _p416;
(* Rung 278 *)
_p417 := Output_Share_M[4] AND TimerQ_In_SenCY_Sep_Claw1_F AND TimerQ_In_SenCY_Sep_Claw2_F;
Out_CYw_Sep_Claw_F_Done := _p417;
Output_Share_Reset_TON[4](In := _p417, PT := T#1s);
(* Rung 279: 異常監視（自動指令・到達待ち10秒） *)
Output_Share_Error_TON[4](In := Out_CYw_Sep_Claw_F_Auto[1] AND AutoMode AND NOT Pause[1] AND ((NOT TimerQ_In_SenCY_Sep_Claw1_F AND NOT TimerQ_In_SenCY_Sep_Claw2_F) OR (TimerQ_In_SenCY_Sep_Claw1_F AND NOT TimerQ_In_SenCY_Sep_Claw2_F) OR (NOT TimerQ_In_SenCY_Sep_Claw1_F AND TimerQ_In_SenCY_Sep_Claw2_F)), PT := T#10s);
_e418(CLK := Output_Share_Error_TON[4].Q);
IF _e418.Q THEN Output_Share_Error_M[4] := TRUE; END_IF;
HMI_Message_Request[88] := _e418.Q;

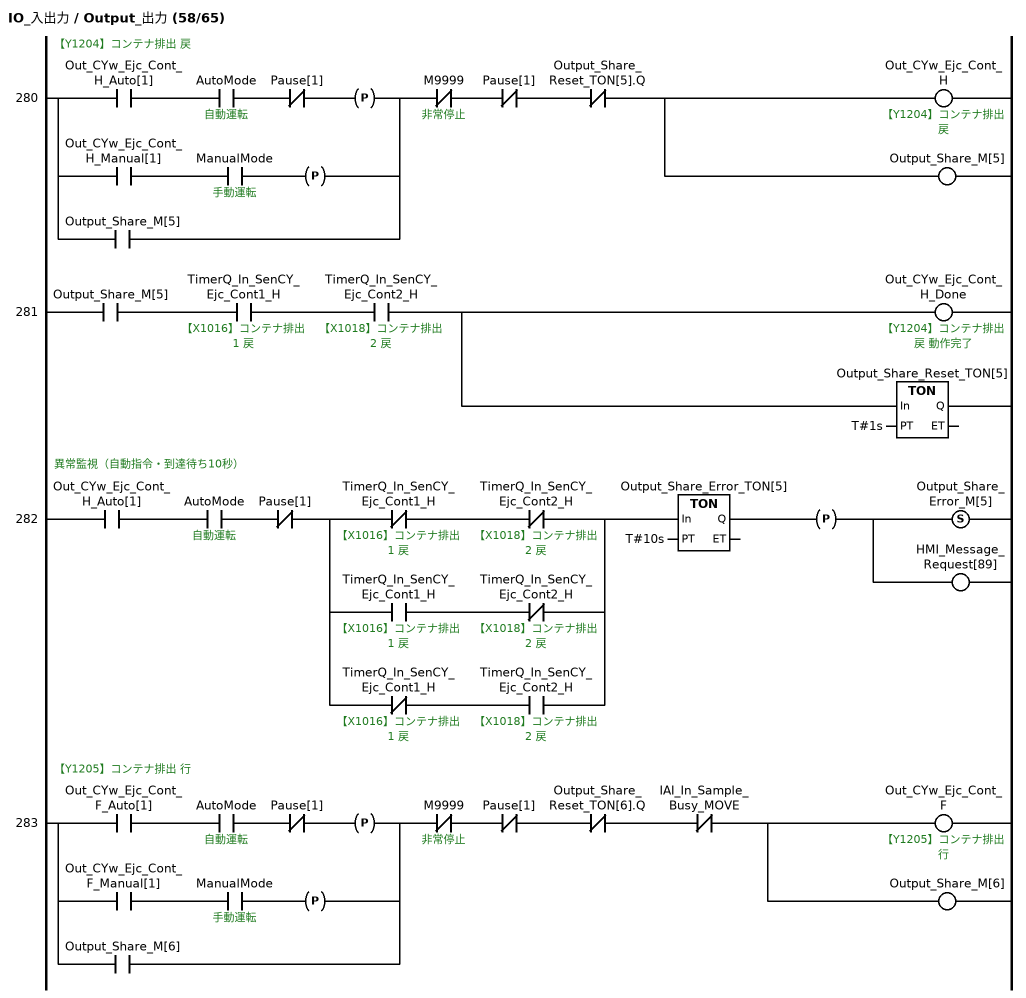
(* Rung 280: 【Y1204】コンテナ排出 戻 *)
_e419(CLK := Out_CYw_Ejc_Cont_H_Auto[1] AND AutoMode AND NOT Pause[1]);
_e420(CLK := Out_CYw_Ejc_Cont_H_Manual[1] AND ManualMode);
_p421 := (_e419.Q OR _e420.Q OR Output_Share_M[5]) AND NOT M9999 AND NOT Pause[1] AND NOT Output_Share_Reset_TON[5].Q;
Out_CYw_Ejc_Cont_H := _p421;
Output_Share_M[5] := _p421;
(* Rung 281 *)
_p422 := Output_Share_M[5] AND TimerQ_In_SenCY_Ejc_Cont1_H AND TimerQ_In_SenCY_Ejc_Cont2_H;
Out_CYw_Ejc_Cont_H_Done := _p422;
Output_Share_Reset_TON[5](In := _p422, PT := T#1s);
(* Rung 282: 異常監視（自動指令・到達待ち10秒） *)
Output_Share_Error_TON[5](In := Out_CYw_Ejc_Cont_H_Auto[1] AND AutoMode AND NOT Pause[1] AND ((NOT TimerQ_In_SenCY_Ejc_Cont1_H AND NOT TimerQ_In_SenCY_Ejc_Cont2_H) OR (TimerQ_In_SenCY_Ejc_Cont1_H AND NOT TimerQ_In_SenCY_Ejc_Cont2_H) OR (NOT TimerQ_In_SenCY_Ejc_Cont1_H AND TimerQ_In_SenCY_Ejc_Cont2_H)), PT := T#10s);
_e423(CLK := Output_Share_Error_TON[5].Q);
IF _e423.Q THEN Output_Share_Error_M[5] := TRUE; END_IF;
HMI_Message_Request[89] := _e423.Q;
(* Rung 283: 【Y1205】コンテナ排出 行 *)
_e424(CLK := Out_CYw_Ejc_Cont_F_Auto[1] AND AutoMode AND NOT Pause[1]);
_e425(CLK := Out_CYw_Ejc_Cont_F_Manual[1] AND ManualMode);
_p426 := (_e424.Q OR _e425.Q OR Output_Share_M[6]) AND NOT M9999 AND NOT Pause[1] AND NOT Output_Share_Reset_TON[6].Q AND NOT IAI_In_Sample_Busy_MOVE;
Out_CYw_Ejc_Cont_F := _p426;
Output_Share_M[6] := _p426;

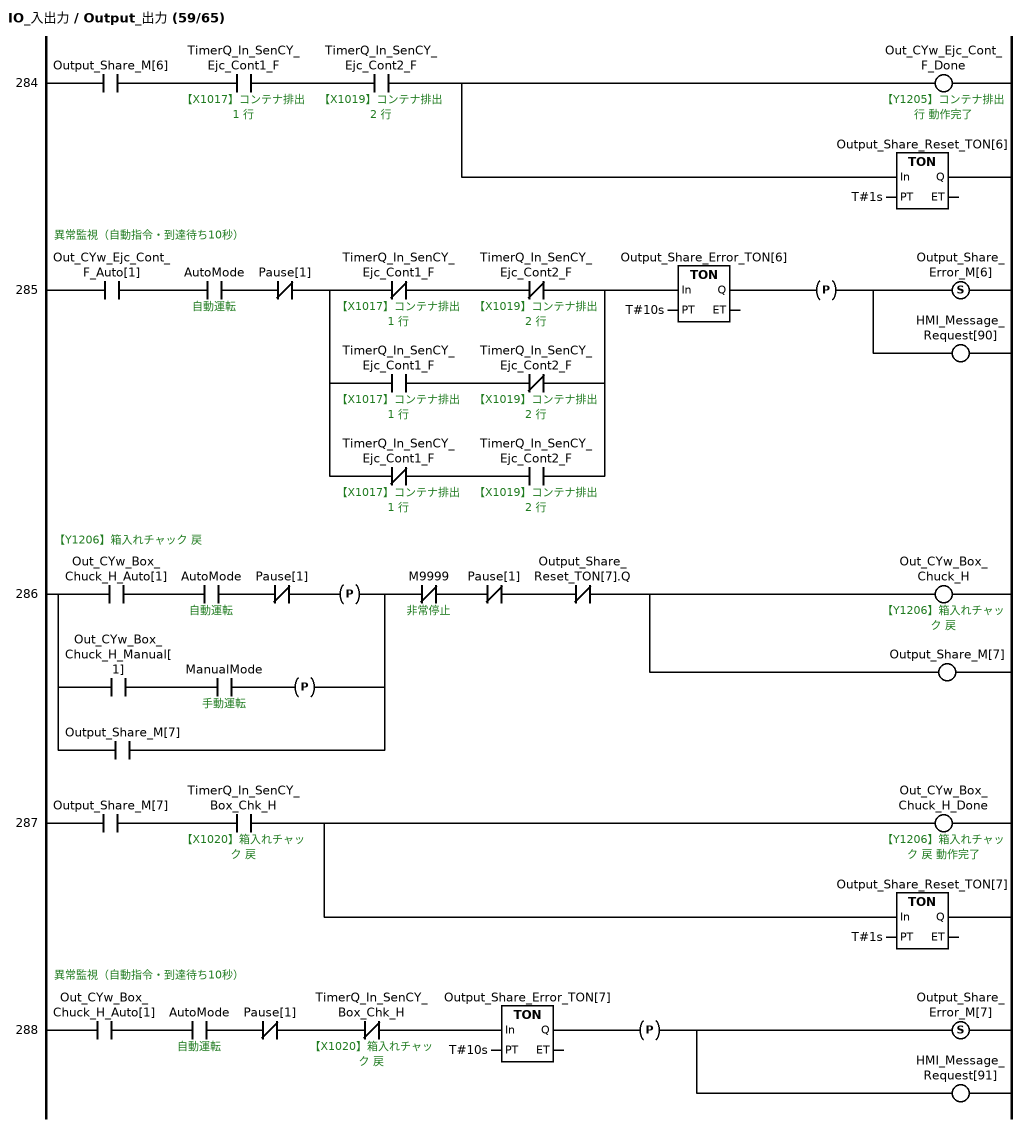
(* Rung 284 *)
_p427 := Output_Share_M[6] AND TimerQ_In_SenCY_Ejc_Cont1_F AND TimerQ_In_SenCY_Ejc_Cont2_F;
Out_CYw_Ejc_Cont_F_Done := _p427;
Output_Share_Reset_TON[6](In := _p427, PT := T#1s);
(* Rung 285: 異常監視（自動指令・到達待ち10秒） *)
Output_Share_Error_TON[6](In := Out_CYw_Ejc_Cont_F_Auto[1] AND AutoMode AND NOT Pause[1] AND ((NOT TimerQ_In_SenCY_Ejc_Cont1_F AND NOT TimerQ_In_SenCY_Ejc_Cont2_F) OR (TimerQ_In_SenCY_Ejc_Cont1_F AND NOT TimerQ_In_SenCY_Ejc_Cont2_F) OR (NOT TimerQ_In_SenCY_Ejc_Cont1_F AND TimerQ_In_SenCY_Ejc_Cont2_F)), PT := T#10s);
_e428(CLK := Output_Share_Error_TON[6].Q);
IF _e428.Q THEN Output_Share_Error_M[6] := TRUE; END_IF;
HMI_Message_Request[90] := _e428.Q;
(* Rung 286: 【Y1206】箱入れチャック 戻 *)
_e429(CLK := Out_CYw_Box_Chuck_H_Auto[1] AND AutoMode AND NOT Pause[1]);
_e430(CLK := Out_CYw_Box_Chuck_H_Manual[1] AND ManualMode);
_p431 := (_e429.Q OR _e430.Q OR Output_Share_M[7]) AND NOT M9999 AND NOT Pause[1] AND NOT Output_Share_Reset_TON[7].Q;
Out_CYw_Box_Chuck_H := _p431;
Output_Share_M[7] := _p431;
(* Rung 287 *)
Out_CYw_Box_Chuck_H_Done := Output_Share_M[7] AND TimerQ_In_SenCY_Box_Chk_H;
Output_Share_Reset_TON[7](In := Output_Share_M[7] AND TimerQ_In_SenCY_Box_Chk_H, PT := T#1s);
(* Rung 288: 異常監視（自動指令・到達待ち10秒） *)
Output_Share_Error_TON[7](In := Out_CYw_Box_Chuck_H_Auto[1] AND AutoMode AND NOT Pause[1] AND NOT TimerQ_In_SenCY_Box_Chk_H, PT := T#10s);
_e432(CLK := Output_Share_Error_TON[7].Q);
IF _e432.Q THEN Output_Share_Error_M[7] := TRUE; END_IF;
HMI_Message_Request[91] := _e432.Q;

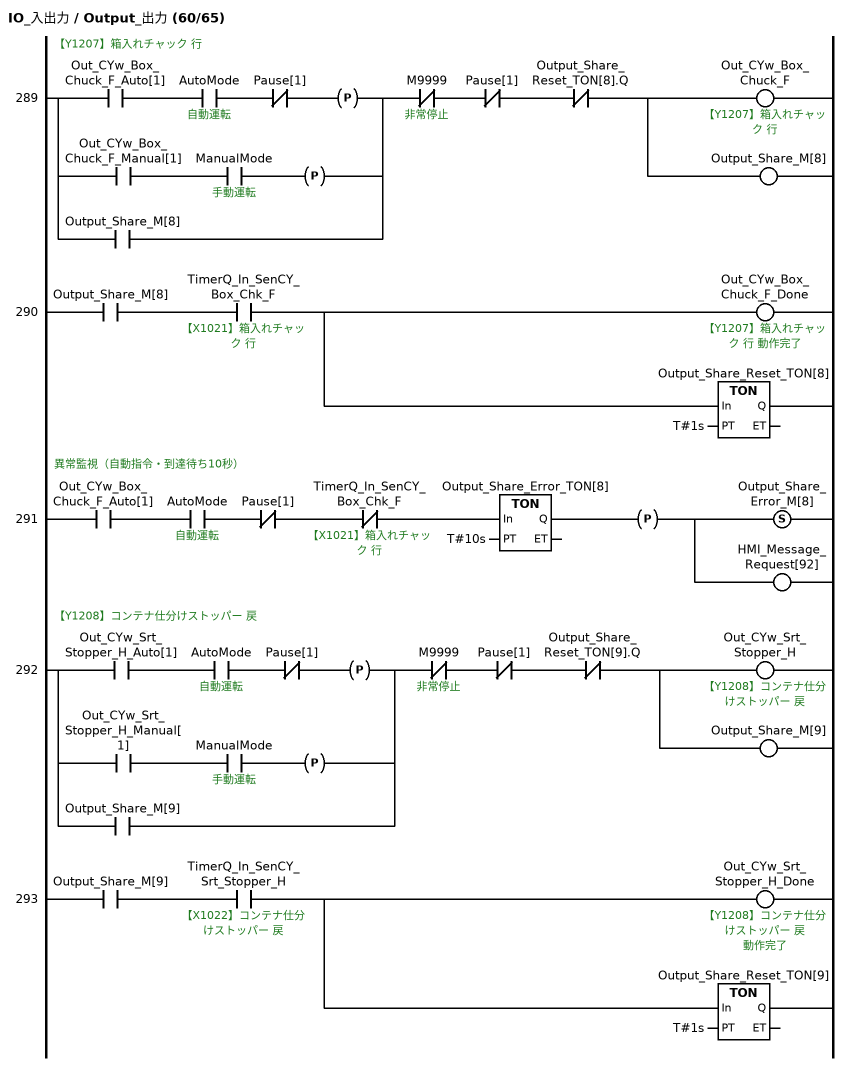
(* Rung 289: 【Y1207】箱入れチャック 行 *)
_e433(CLK := Out_CYw_Box_Chuck_F_Auto[1] AND AutoMode AND NOT Pause[1]);
_e434(CLK := Out_CYw_Box_Chuck_F_Manual[1] AND ManualMode);
_p435 := (_e433.Q OR _e434.Q OR Output_Share_M[8]) AND NOT M9999 AND NOT Pause[1] AND NOT Output_Share_Reset_TON[8].Q;
Out_CYw_Box_Chuck_F := _p435;
Output_Share_M[8] := _p435;
(* Rung 290 *)
Out_CYw_Box_Chuck_F_Done := Output_Share_M[8] AND TimerQ_In_SenCY_Box_Chk_F;
Output_Share_Reset_TON[8](In := Output_Share_M[8] AND TimerQ_In_SenCY_Box_Chk_F, PT := T#1s);
(* Rung 291: 異常監視（自動指令・到達待ち10秒） *)
Output_Share_Error_TON[8](In := Out_CYw_Box_Chuck_F_Auto[1] AND AutoMode AND NOT Pause[1] AND NOT TimerQ_In_SenCY_Box_Chk_F, PT := T#10s);
_e436(CLK := Output_Share_Error_TON[8].Q);
IF _e436.Q THEN Output_Share_Error_M[8] := TRUE; END_IF;
HMI_Message_Request[92] := _e436.Q;
(* Rung 292: 【Y1208】コンテナ仕分けストッパー 戻 *)
_e437(CLK := Out_CYw_Srt_Stopper_H_Auto[1] AND AutoMode AND NOT Pause[1]);
_e438(CLK := Out_CYw_Srt_Stopper_H_Manual[1] AND ManualMode);
_p439 := (_e437.Q OR _e438.Q OR Output_Share_M[9]) AND NOT M9999 AND NOT Pause[1] AND NOT Output_Share_Reset_TON[9].Q;
Out_CYw_Srt_Stopper_H := _p439;
Output_Share_M[9] := _p439;
(* Rung 293 *)
_p440 := Output_Share_M[9] AND TimerQ_In_SenCY_Srt_Stopper_H;
Out_CYw_Srt_Stopper_H_Done := _p440;
Output_Share_Reset_TON[9](In := _p440, PT := T#1s);

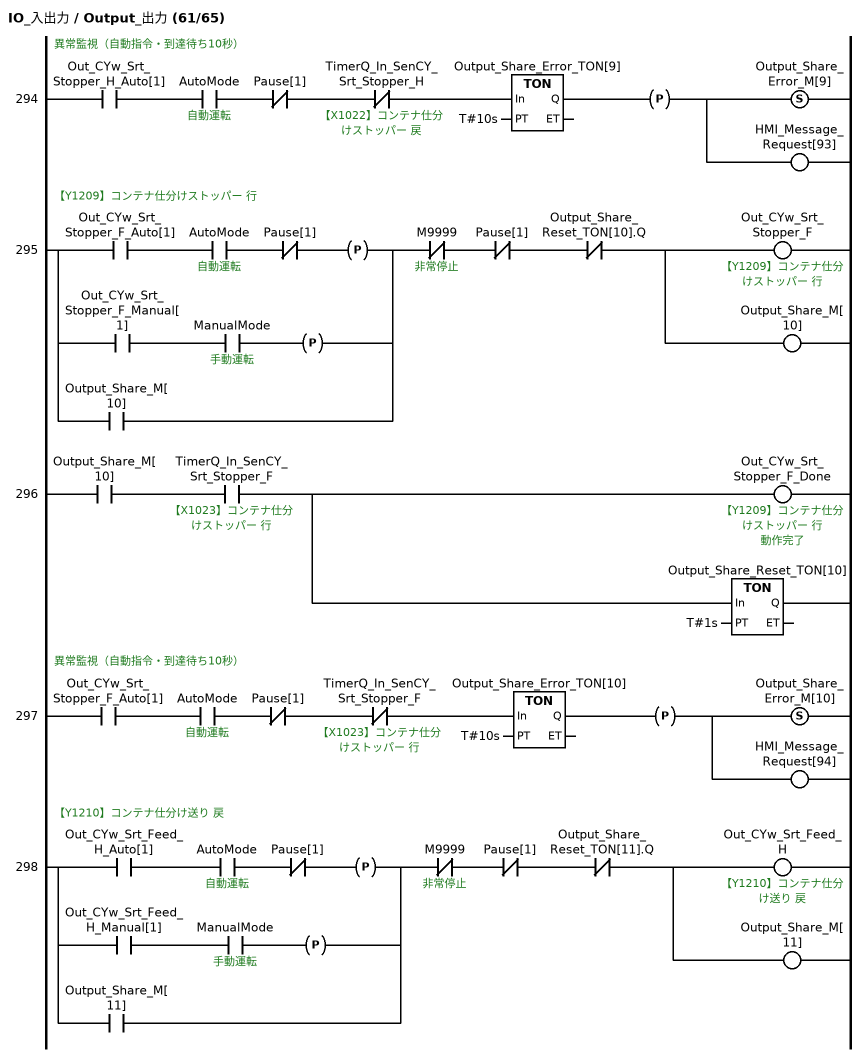
(* Rung 294: 異常監視（自動指令・到達待ち10秒） *)
Output_Share_Error_TON[9](In := Out_CYw_Srt_Stopper_H_Auto[1] AND AutoMode AND NOT Pause[1] AND NOT TimerQ_In_SenCY_Srt_Stopper_H, PT := T#10s);
_e441(CLK := Output_Share_Error_TON[9].Q);
IF _e441.Q THEN Output_Share_Error_M[9] := TRUE; END_IF;
HMI_Message_Request[93] := _e441.Q;
(* Rung 295: 【Y1209】コンテナ仕分けストッパー 行 *)
_e442(CLK := Out_CYw_Srt_Stopper_F_Auto[1] AND AutoMode AND NOT Pause[1]);
_e443(CLK := Out_CYw_Srt_Stopper_F_Manual[1] AND ManualMode);
_p444 := (_e442.Q OR _e443.Q OR Output_Share_M[10]) AND NOT M9999 AND NOT Pause[1] AND NOT Output_Share_Reset_TON[10].Q;
Out_CYw_Srt_Stopper_F := _p444;
Output_Share_M[10] := _p444;
(* Rung 296 *)
_p445 := Output_Share_M[10] AND TimerQ_In_SenCY_Srt_Stopper_F;
Out_CYw_Srt_Stopper_F_Done := _p445;
Output_Share_Reset_TON[10](In := _p445, PT := T#1s);
(* Rung 297: 異常監視（自動指令・到達待ち10秒） *)
Output_Share_Error_TON[10](In := Out_CYw_Srt_Stopper_F_Auto[1] AND AutoMode AND NOT Pause[1] AND NOT TimerQ_In_SenCY_Srt_Stopper_F, PT := T#10s);
_e446(CLK := Output_Share_Error_TON[10].Q);
IF _e446.Q THEN Output_Share_Error_M[10] := TRUE; END_IF;
HMI_Message_Request[94] := _e446.Q;
(* Rung 298: 【Y1210】コンテナ仕分け送り 戻 *)
_e447(CLK := Out_CYw_Srt_Feed_H_Auto[1] AND AutoMode AND NOT Pause[1]);
_e448(CLK := Out_CYw_Srt_Feed_H_Manual[1] AND ManualMode);
_p449 := (_e447.Q OR _e448.Q OR Output_Share_M[11]) AND NOT M9999 AND NOT Pause[1] AND NOT Output_Share_Reset_TON[11].Q;
Out_CYw_Srt_Feed_H := _p449;
Output_Share_M[11] := _p449;

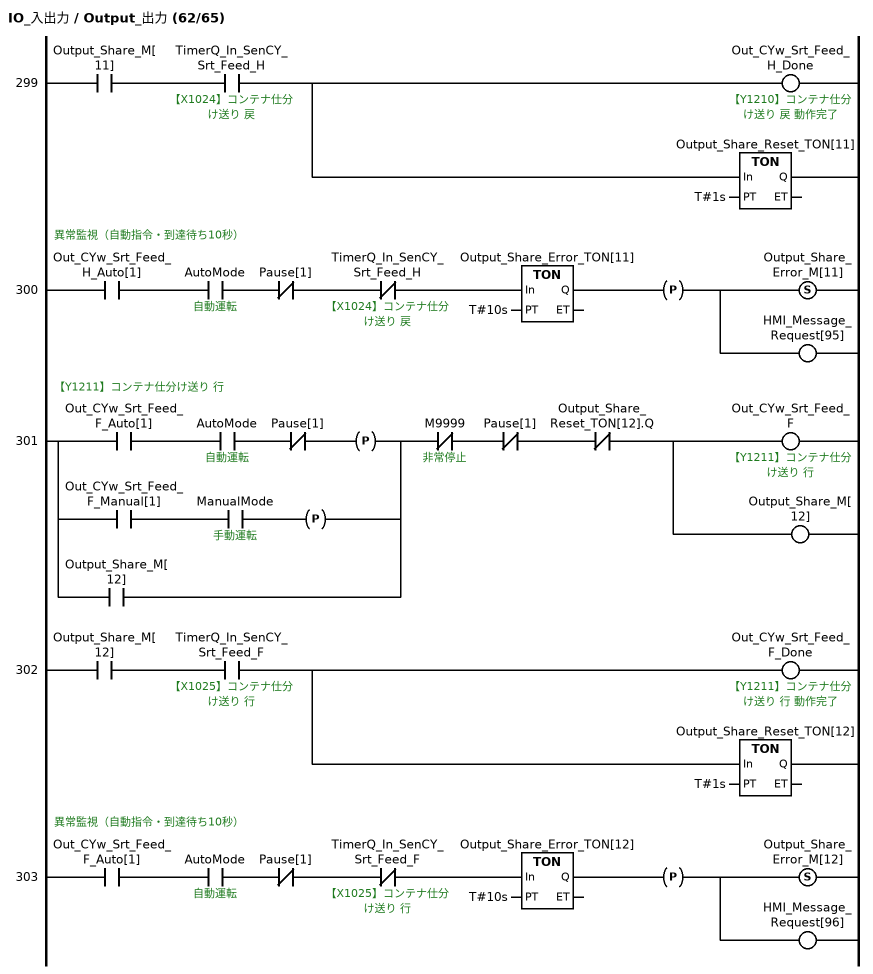
(* Rung 299 *)
_p450 := Output_Share_M[11] AND TimerQ_In_SenCY_Srt_Feed_H;
Out_CYw_Srt_Feed_H_Done := _p450;
Output_Share_Reset_TON[11](In := _p450, PT := T#1s);
(* Rung 300: 異常監視（自動指令・到達待ち10秒） *)
Output_Share_Error_TON[11](In := Out_CYw_Srt_Feed_H_Auto[1] AND AutoMode AND NOT Pause[1] AND NOT TimerQ_In_SenCY_Srt_Feed_H, PT := T#10s);
_e451(CLK := Output_Share_Error_TON[11].Q);
IF _e451.Q THEN Output_Share_Error_M[11] := TRUE; END_IF;
HMI_Message_Request[95] := _e451.Q;
(* Rung 301: 【Y1211】コンテナ仕分け送り 行 *)
_e452(CLK := Out_CYw_Srt_Feed_F_Auto[1] AND AutoMode AND NOT Pause[1]);
_e453(CLK := Out_CYw_Srt_Feed_F_Manual[1] AND ManualMode);
_p454 := (_e452.Q OR _e453.Q OR Output_Share_M[12]) AND NOT M9999 AND NOT Pause[1] AND NOT Output_Share_Reset_TON[12].Q;
Out_CYw_Srt_Feed_F := _p454;
Output_Share_M[12] := _p454;
(* Rung 302 *)
_p455 := Output_Share_M[12] AND TimerQ_In_SenCY_Srt_Feed_F;
Out_CYw_Srt_Feed_F_Done := _p455;
Output_Share_Reset_TON[12](In := _p455, PT := T#1s);
(* Rung 303: 異常監視（自動指令・到達待ち10秒） *)
Output_Share_Error_TON[12](In := Out_CYw_Srt_Feed_F_Auto[1] AND AutoMode AND NOT Pause[1] AND NOT TimerQ_In_SenCY_Srt_Feed_F, PT := T#10s);
_e456(CLK := Output_Share_Error_TON[12].Q);
IF _e456.Q THEN Output_Share_Error_M[12] := TRUE; END_IF;
HMI_Message_Request[96] := _e456.Q;

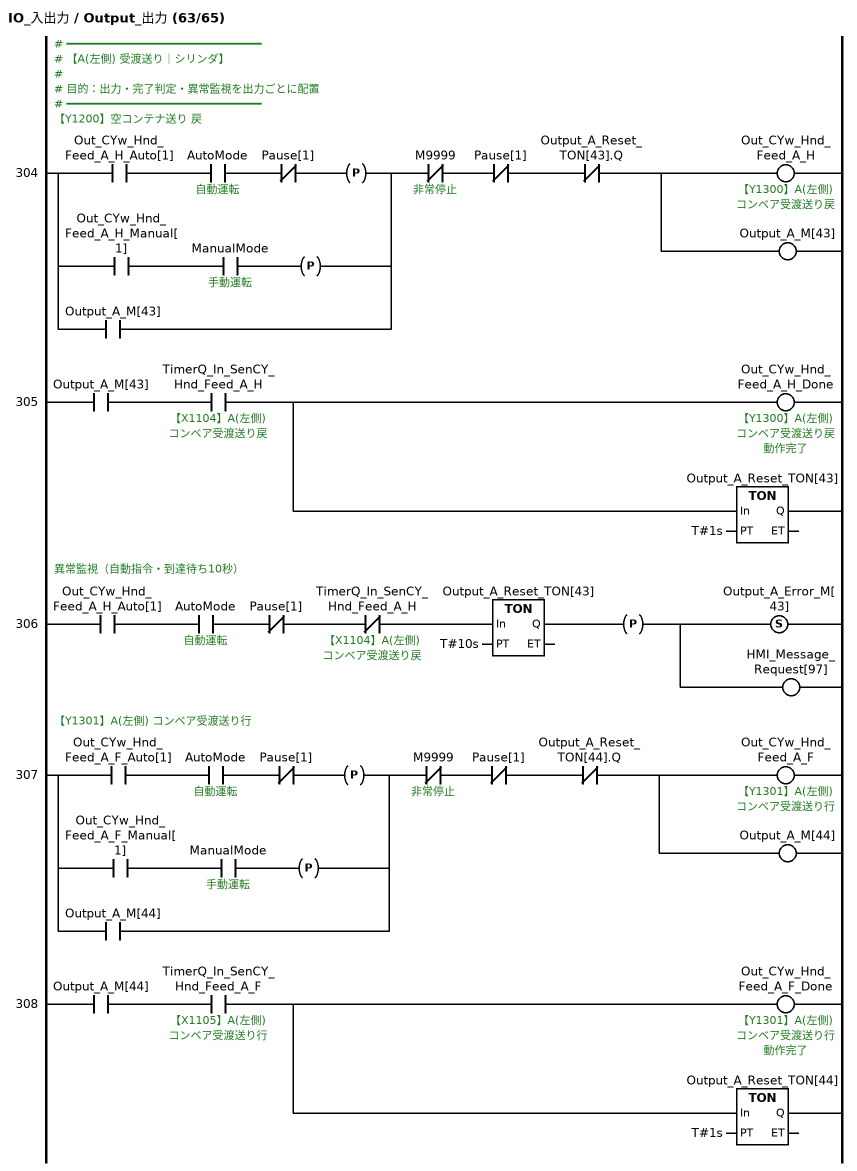
(* Rung 304: # ━━━━━━━━━━━━━━━━━━━━━━━━━━━━━━ / # 【A(左側) 受渡送り｜シリンダ】 / # / # 目的：出力・完了判定・異常監視を出力ごとに配置 / # ━━━━━━━━━━━━━━━━━━━━━━━━━━━━━━ / 【Y1200】空コンテナ送り 戻 *)
_e457(CLK := Out_CYw_Hnd_Feed_A_H_Auto[1] AND AutoMode AND NOT Pause[1]);
_e458(CLK := Out_CYw_Hnd_Feed_A_H_Manual[1] AND ManualMode);
_p459 := (_e457.Q OR _e458.Q OR Output_A_M[43]) AND NOT M9999 AND NOT Pause[1] AND NOT Output_A_Reset_TON[43].Q;
Out_CYw_Hnd_Feed_A_H := _p459;
Output_A_M[43] := _p459;
(* Rung 305 *)
Out_CYw_Hnd_Feed_A_H_Done := Output_A_M[43] AND TimerQ_In_SenCY_Hnd_Feed_A_H;
Output_A_Reset_TON[43](In := Output_A_M[43] AND TimerQ_In_SenCY_Hnd_Feed_A_H, PT := T#1s);
(* Rung 306: 異常監視（自動指令・到達待ち10秒） *)
Output_A_Reset_TON[43](In := Out_CYw_Hnd_Feed_A_H_Auto[1] AND AutoMode AND NOT Pause[1] AND NOT TimerQ_In_SenCY_Hnd_Feed_A_H, PT := T#10s);
_e460(CLK := Output_A_Reset_TON[43].Q);
IF _e460.Q THEN Output_A_Error_M[43] := TRUE; END_IF;
HMI_Message_Request[97] := _e460.Q;
(* Rung 307: 【Y1301】A(左側) コンベア受渡送り行 *)
_e461(CLK := Out_CYw_Hnd_Feed_A_F_Auto[1] AND AutoMode AND NOT Pause[1]);
_e462(CLK := Out_CYw_Hnd_Feed_A_F_Manual[1] AND ManualMode);
_p463 := (_e461.Q OR _e462.Q OR Output_A_M[44]) AND NOT M9999 AND NOT Pause[1] AND NOT Output_A_Reset_TON[44].Q;
Out_CYw_Hnd_Feed_A_F := _p463;
Output_A_M[44] := _p463;
(* Rung 308 *)
Out_CYw_Hnd_Feed_A_F_Done := Output_A_M[44] AND TimerQ_In_SenCY_Hnd_Feed_A_F;
Output_A_Reset_TON[44](In := Output_A_M[44] AND TimerQ_In_SenCY_Hnd_Feed_A_F, PT := T#1s);

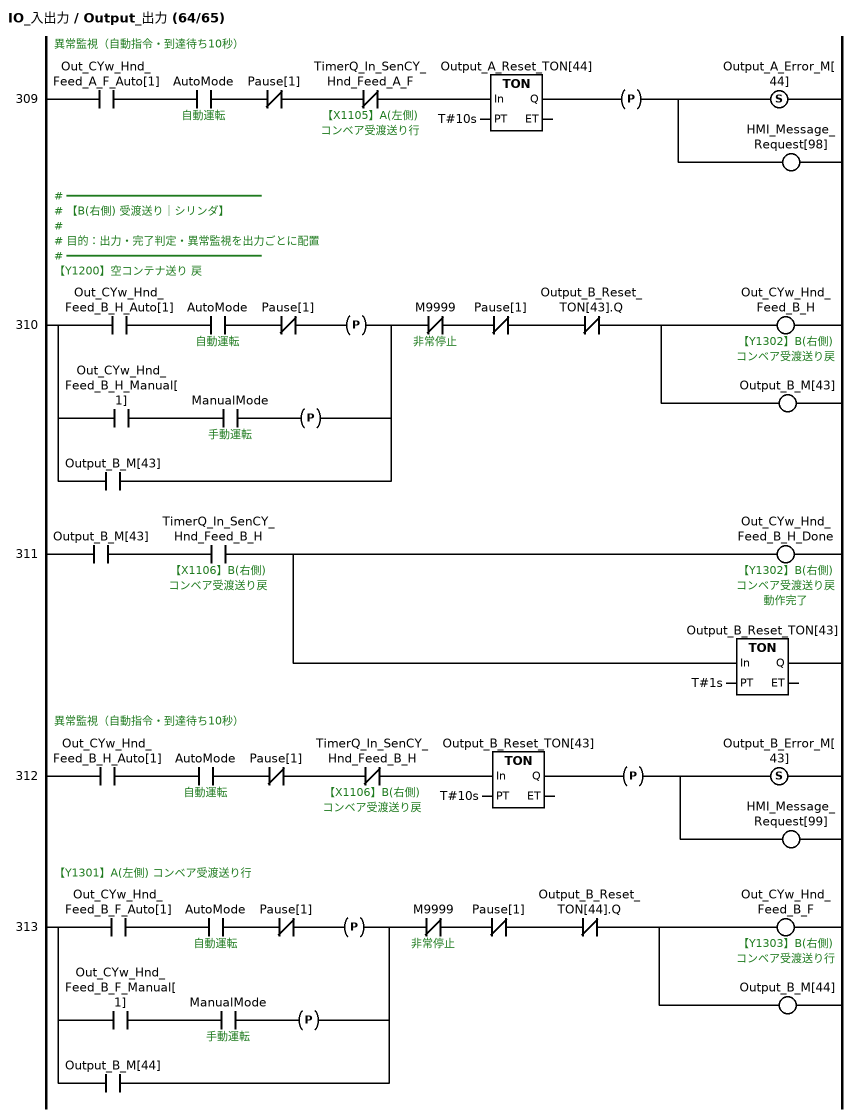
(* Rung 309: 異常監視（自動指令・到達待ち10秒） *)
Output_A_Reset_TON[44](In := Out_CYw_Hnd_Feed_A_F_Auto[1] AND AutoMode AND NOT Pause[1] AND NOT TimerQ_In_SenCY_Hnd_Feed_A_F, PT := T#10s);
_e464(CLK := Output_A_Reset_TON[44].Q);
IF _e464.Q THEN Output_A_Error_M[44] := TRUE; END_IF;
HMI_Message_Request[98] := _e464.Q;
(* Rung 310: # ━━━━━━━━━━━━━━━━━━━━━━━━━━━━━━ / # 【B(右側) 受渡送り｜シリンダ】 / # / # 目的：出力・完了判定・異常監視を出力ごとに配置 / # ━━━━━━━━━━━━━━━━━━━━━━━━━━━━━━ / 【Y1200】空コンテナ送り 戻 *)
_e465(CLK := Out_CYw_Hnd_Feed_B_H_Auto[1] AND AutoMode AND NOT Pause[1]);
_e466(CLK := Out_CYw_Hnd_Feed_B_H_Manual[1] AND ManualMode);
_p467 := (_e465.Q OR _e466.Q OR Output_B_M[43]) AND NOT M9999 AND NOT Pause[1] AND NOT Output_B_Reset_TON[43].Q;
Out_CYw_Hnd_Feed_B_H := _p467;
Output_B_M[43] := _p467;
(* Rung 311 *)
Out_CYw_Hnd_Feed_B_H_Done := Output_B_M[43] AND TimerQ_In_SenCY_Hnd_Feed_B_H;
Output_B_Reset_TON[43](In := Output_B_M[43] AND TimerQ_In_SenCY_Hnd_Feed_B_H, PT := T#1s);
(* Rung 312: 異常監視（自動指令・到達待ち10秒） *)
Output_B_Reset_TON[43](In := Out_CYw_Hnd_Feed_B_H_Auto[1] AND AutoMode AND NOT Pause[1] AND NOT TimerQ_In_SenCY_Hnd_Feed_B_H, PT := T#10s);
_e468(CLK := Output_B_Reset_TON[43].Q);
IF _e468.Q THEN Output_B_Error_M[43] := TRUE; END_IF;
HMI_Message_Request[99] := _e468.Q;
(* Rung 313: 【Y1301】A(左側) コンベア受渡送り行 *)
_e469(CLK := Out_CYw_Hnd_Feed_B_F_Auto[1] AND AutoMode AND NOT Pause[1]);
_e470(CLK := Out_CYw_Hnd_Feed_B_F_Manual[1] AND ManualMode);
_p471 := (_e469.Q OR _e470.Q OR Output_B_M[44]) AND NOT M9999 AND NOT Pause[1] AND NOT Output_B_Reset_TON[44].Q;
Out_CYw_Hnd_Feed_B_F := _p471;
Output_B_M[44] := _p471;

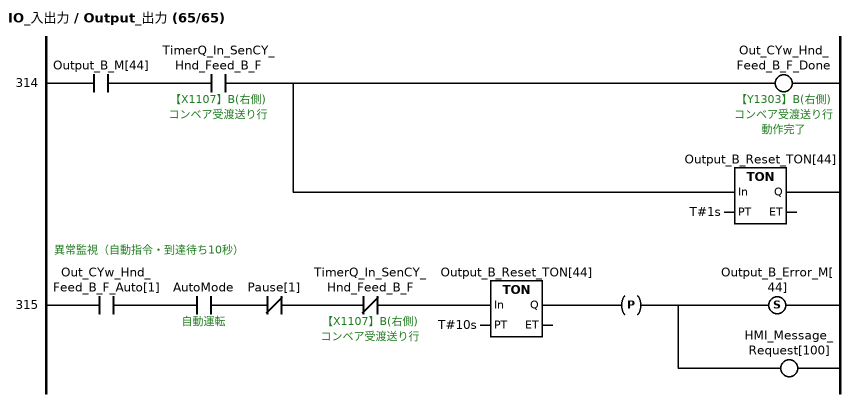
(* Rung 314 *)
Out_CYw_Hnd_Feed_B_F_Done := Output_B_M[44] AND TimerQ_In_SenCY_Hnd_Feed_B_F;
Output_B_Reset_TON[44](In := Output_B_M[44] AND TimerQ_In_SenCY_Hnd_Feed_B_F, PT := T#1s);
(* Rung 315: 異常監視（自動指令・到達待ち10秒） *)
Output_B_Reset_TON[44](In := Out_CYw_Hnd_Feed_B_F_Auto[1] AND AutoMode AND NOT Pause[1] AND NOT TimerQ_In_SenCY_Hnd_Feed_B_F, PT := T#10s);
_e472(CLK := Output_B_Reset_TON[44].Q);
IF _e472.Q THEN Output_B_Error_M[44] := TRUE; END_IF;
HMI_Message_Request[100] := _e472.Q;
END_PROGRAM

# Device HMI_NA5_0 (NA): not converted